(* IEC 61131-3 sources: daoli-st-library/DL_Process (part 19) *)

(* ---- FC_DL_WeighSpanCalibRatio.st ---- *)
(*
  ============================================================
  组件名 : FC_DL_WeighSpanCalibRatio
  分类   : DL_Process
  功能   : 称重系统量程标定，由零点和量程两点原始值求比例系数与量程误差
  开源溯源 : internal-design（本轮无外部代码逐行引用）
             参考语义 : 无外部参考
  复杂度 : C1
  版本   : 1.0.0
  ============================================================
*)

FUNCTION FC_DL_WeighSpanCalibRatio : REAL
VAR_INPUT
    rRawAtZero : REAL; // 空载时原始值 [count] raw value at no load [count]
    rRawAtSpan : REAL; // 加载标准砝码时原始值 [count] raw value at the reference span [count]
    rRefSpan   : REAL; // 标准砝码标称值 [kg] nominal reference weight [kg]
END_VAR
VAR_OUTPUT
    rRatio        : REAL; // 标定比例系数 [kg/count] calibration ratio [kg per count]
    rSpanErrorPct : REAL; // 量程误差百分比 [%] span error percentage [%]
    bValid        : BOOL; // 结果有效标志 result validity flag
END_VAR
VAR CONSTANT
    DL_EPS_R    : REAL := 1.0E-6; // 实数零判定阈值 real zero threshold
    DL_ERR_LIM  : REAL := 5.0; // 量程误差合理上限 [%] admissible span error ceiling [%]
    DL_HUNDRED  : REAL := 100.0; // 百分制换算系数 percentage scale factor
END_VAR
VAR
    _bFin   : BOOL := FALSE; // 三输入有限性判定 finiteness verdict of the three inputs
    _rDelta : REAL := 0.0; // 两点原始值增量 [count] raw span increment [count]
    _rRatio : REAL := 0.0; // 比例系数中间量 [kg/count] intermediate ratio [kg per count]
    _rErr   : REAL := 0.0; // 量程误差中间量 [%] intermediate span error [%]
    _rPred  : REAL := 0.0; // 按比例反推的砝码值 [kg] weight predicted by the ratio [kg]
END_VAR

// 段 1｜出口预置 preset the exit
FC_DL_WeighSpanCalibRatio := 0.0; // 缺省返回零 default zero return
rRatio := 0.0; // 比例系数预置零 ratio preset to zero
rSpanErrorPct := 0.0; // 量程误差预置零 span error preset to zero
bValid := FALSE; // 计算完成前不认结果 unusable before the calculation
// 段 2｜非有限闸 finiteness gate
_bFin := (rRawAtZero = rRawAtZero) AND (rRawAtSpan = rRawAtSpan) AND (rRefSpan = rRefSpan); // 三输入自反判定 self comparison of the three inputs
IF NOT _bFin THEN
    RETURN; // 非有限即无效 non finite means invalid
END_IF
// 段 3｜两点增量与砝码值闸 span increment and reference weight gate
_rDelta := rRawAtSpan - rRawAtZero; // 量程段原始增量 raw increment over the span
IF (ABS(_rDelta) < DL_EPS_R) OR (rRefSpan <= 0.0) THEN
    RETURN; // 增量近零或砝码非正无法标定 a zero increment or a non positive reference cannot calibrate
END_IF
// 段 4｜比例系数与量程误差 ratio and span error
_rRatio := rRefSpan / _rDelta; // 比例系数 ratio of the reference to the increment
_rPred := _rRatio * rRefSpan; // 按比例反推的砝码值 weight predicted from the ratio
_rErr := (_rPred - rRefSpan) / rRefSpan * DL_HUNDRED; // 量程误差百分比 span error percentage
rRatio := _rRatio; // 比例系数落定 land the ratio
rSpanErrorPct := _rErr; // 量程误差落定 land the span error
// 段 5｜超差合理性闸 span error plausibility gate
IF ABS(_rErr) > DL_ERR_LIM THEN
    RETURN; // 超差判无效，比例系数保留供诊断 an excessive error is void while the ratio stays for diagnosis
END_IF
bValid := TRUE; // 结果可用 result usable
FC_DL_WeighSpanCalibRatio := _rRatio; // 函数返回比例系数 return the ratio
END_FUNCTION

(* ---- FC_DL_WeighTareDriftCheck.st ---- *)
(*
  ============================================================
  组件名 : FC_DL_WeighTareDriftCheck
  分类   : DL_Process
  功能   : 单点皮重相对标定基准的漂移量与漂移百分比监视，超限置位
  开源溯源 : internal-design（本轮无外部代码逐行引用）
             参考语义 : 无外部参考
  复杂度 : C1
  版本   : 1.0.0
  ============================================================
*)

FUNCTION FC_DL_WeighTareDriftCheck : BOOL
VAR_INPUT
    rTareNow    : REAL; // 当前实测皮重 [kg] current measured tare [kg]
    rTareRef    : REAL; // 标定基准皮重 [kg] calibrated reference tare [kg]
    rDriftLimit : REAL; // 漂移报警限 [kg] drift alarm limit [kg]
    nSamples    : INT; // 采样点数 [个] sample count [count]
END_VAR
VAR_OUTPUT
    rDrift         : REAL; // 皮重漂移量 [kg] tare drift [kg]
    rDriftPct      : REAL; // 漂移百分比 [%] drift percentage [%]
    bDriftExceeded : BOOL; // 漂移超限标志 drift exceeded flag
    bValid         : BOOL; // 结果有效标志 result validity flag
END_VAR
VAR CONSTANT
    DL_EPS_R : REAL := 1.0E-6; // 实数零判定阈值 real zero threshold
END_VAR
VAR
    _bFin : BOOL := FALSE; // 三实数输入有限性判定 finiteness verdict of the three real inputs
    _rLim : REAL := 0.0; // 钳位后的漂移限 [kg] clamped drift limit [kg]
END_VAR

// 段 1｜出口预置 preset the exit
FC_DL_WeighTareDriftCheck := FALSE; // 缺省返回未超限 default not exceeded
rDrift := 0.0; // 漂移量预置零 drift preset to zero
rDriftPct := 0.0; // 漂移百分比预置零 drift percentage preset to zero
bDriftExceeded := FALSE; // 超限标志预置假 exceeded flag preset false
bValid := FALSE; // 计算完成前不认结果 unusable before the calculation
// 段 2｜非有限闸与点数闸 finiteness gate and sample count gate
_bFin := (rTareNow = rTareNow) AND (rTareRef = rTareRef) AND (rDriftLimit = rDriftLimit); // 三输入自反判定 self comparison of the three inputs
IF (NOT _bFin) OR (nSamples < 1) THEN
    RETURN; // 非有限或无采样即无效 non finite or no sample means invalid
END_IF
// 段 3｜漂移量与百分比 drift value and percentage
rDrift := rTareNow - rTareRef; // 单点滑动漂移量 single point sliding drift
IF ABS(rTareRef) < DL_EPS_R THEN
    RETURN; // 基准皮重近零无法折算百分比 a zero reference cannot carry a percentage
END_IF
rDriftPct := rDrift / rTareRef * 100.0; // 相对基准的漂移百分比 drift relative to the reference [%]
// 段 4｜限值整形与超限判定 limit reshape and the exceed verdict
_rLim := rDriftLimit; // 取入参限值 take the limit input
IF _rLim < 0.0 THEN
    _rLim := ABS(_rLim); // 负限值取幅值 a negative limit becomes its magnitude
END_IF
bDriftExceeded := ABS(rDrift) > _rLim; // 双向漂移均计入超限 drift counts in both directions
bValid := TRUE; // 结果可用 result usable
FC_DL_WeighTareDriftCheck := bDriftExceeded; // 函数返回超限标志 return the exceeded flag
END_FUNCTION

(* ---- FC_DL_WortAerationRateCalc.st ---- *)
// FC_DL_WortAerationRateCalc v1.0.0
// 开源溯源：clean-room 自研（族 DL_Process，ST 生态实测 0 命中，无外部代码引入）
(*
  功能: 麦汁溶解氧：供氧质量 = 风量·1.429·氧体积分数·吸收效率 [kg/h]（1.429 为标况氧密度），
        麦汁体积 = 流量[hL/h]·100 [L/h]，溶解氧 = 供氧/体积 [g/L]→×1000 [mg/L]（等值 ppm）。
  邻件/码位: 位于煮沸之后、接种之前；与 FC_DL_YeastPitchRateCalc 的接种量直接相关；
             16#0002_9232 = 非有限、麦汁流量非正、空气流量为负、效率或氧分数越界、氧超 20 mg/L。
*)
FUNCTION FC_DL_WortAerationRateCalc : REAL
VAR_INPUT
    fWortFlow  : REAL := 200.0;     // 麦汁流量 [hL/h]，域 > 0 / Wort flow [hL/h]
    fAirFlow   : REAL := 1.71;      // 无菌空气流量 [Nm³/h]，域 >= 0（缺省 1.71 → 约 9.0 mg/L 落 8~10 工艺窗，R92 复裁修）/ Sterile air flow [Nm^3/h]
    fO2Frac    : REAL := 0.21;      // 氧体积分数 [-]，域 (0, 1] / Oxygen fraction
    fAbsorbEff : REAL := 0.35;      // 吸收效率 [-]，域 (0, 1] / Absorption efficiency
END_VAR
VAR_OUTPUT
    fO2ppm   : REAL;                // 溶解氧 [mg/L]（等值 ppm）/ Dissolved oxygen [mg/L]
    bValid   : BOOL;                // 结果有效回执 [-] / Result validity receipt
    uErrorId : UDINT;               // 事件码，0 = 无事件 / Event code
END_VAR
VAR
    fVolLh : REAL := 0.0;           // 麦汁体积流量 [L/h] / Wort volume flow [L/h]
END_VAR
// 段 0：全路径出口安全缺省 / Safe defaults on all outlets
fO2ppm := 0.0;                      // 溶解氧缺省零 / Dissolved oxygen default zero
bValid := FALSE;                    // 有效回执预清 / Validity preset clear
uErrorId := 16#0000;                // 事件码预清 / Event code preset clear
FC_DL_WortAerationRateCalc := 0.0;  // 返回值缺省零（镜像溶解氧）/ Return default zero
// 段 1：非有限闸（四入参全枚举）/ Non-finite gate over all inputs
IF (fWortFlow <> fWortFlow) OR (fAirFlow <> fAirFlow)
   OR (fO2Frac <> fO2Frac) OR (fAbsorbEff <> fAbsorbEff)
   OR (ABS(fWortFlow) >= 3.0E38) OR (ABS(fAirFlow) >= 3.0E38)
   OR (ABS(fO2Frac) >= 3.0E38) OR (ABS(fAbsorbEff) >= 3.0E38) THEN
    uErrorId := 16#0002_9232;   // 入参非有限拒收 / Non-finite input reject
    RETURN;
END_IF
// 段 2：域闸（麦汁流量正防除零 + 空气非负 + 效率与氧分数区间，R4）/ Domain gate
IF fWortFlow <= 1.0E-6 THEN
    uErrorId := 16#0002_9232;   // 麦汁流量非正 / Non-positive wort flow
    RETURN;
END_IF
IF fAirFlow < 0.0 THEN
    uErrorId := 16#0002_9232;   // 空气流量为负 / Negative air flow
    RETURN;
END_IF
IF (fAbsorbEff <= 0.0) OR (fAbsorbEff > 1.0) THEN
    uErrorId := 16#0002_9232;   // 吸收效率越界 / Absorption efficiency out of range
    RETURN;
END_IF
IF (fO2Frac <= 0.0) OR (fO2Frac > 1.0) THEN
    uErrorId := 16#0002_9232;   // 氧体积分数越界 / Oxygen fraction out of range
    RETURN;
END_IF
// 段 3：主计算（供氧质量 → 麦汁体积 → 溶解氧）/ Main computation
fVolLh := fWortFlow * 100.0;                                    // 麦汁体积 [L/h] / Wort volume flow
fO2ppm := fAirFlow * 1.429 * fO2Frac * fAbsorbEff * 1000.0 / fVolLh * 1000.0;  // [mg/L] / Dissolved oxygen
// 段 4：出口闸（非有限复核 + 20 mg/L 工艺界判定）/ Outlet gate
IF (fO2ppm <> fO2ppm) OR (ABS(fO2ppm) >= 3.0E38) OR (fO2ppm < 0.0) THEN
    fO2ppm := 0.0;              // 复核失败回缺省 / Fallback on recheck failure
    uErrorId := 16#0002_9232;   // 出口复核拒收 / Output recheck reject
    RETURN;
END_IF
IF fO2ppm > 20.0 THEN
    uErrorId := 16#0002_9232;   // 信息级：溶解氧超 20 mg/L / Info: oxygen above bound
    RETURN;                     // bValid 保持 FALSE / Validity stays false
END_IF
bValid := TRUE;                 // 有效回执 / Validity receipt
FC_DL_WortAerationRateCalc := fO2ppm;           // 返回值镜像溶解氧 / Return mirrors oxygen
END_FUNCTION

(* ---- FC_DL_WortBoilEvaporationCalc.st ---- *)
// FC_DL_WortBoilEvaporationCalc v1.0.0
// 开源溯源：clean-room 自研（族 DL_Process，ST 生态实测 0 命中，无外部代码引入）
(*
  功能: 煮沸蒸发：总蒸发率 = 100·(前体积 − 后体积)/前体积 [%]，蒸发强度 = 总蒸发率·60/时长 [%/h]。
        煮沸中体积只减不增，后体积大于前体积直接判数据非法。
  邻件/码位: 位于煮沸工序，是麦汁浓度定标的关键质量指标；与 FC_DL_FermentAttenuationCalc 的原浓耦合；
             16#0002_9233 = 非有限、前体积或时长非正、后体积大于前体积或为负拒收。
*)
FUNCTION FC_DL_WortBoilEvaporationCalc : REAL
VAR_INPUT
    fVolBefore : REAL := 250.0;     // 煮沸前体积 [hL]，域 > 0 / Volume before boil [hL]
    fVolAfter  : REAL := 225.0;     // 煮沸后体积 [hL]，域 <= 前体积 / Volume after boil [hL]
    fBoilMin   : REAL := 60.0;      // 煮沸时长 [min]，域 > 0 / Boil duration [min]
END_VAR
VAR_OUTPUT
    fEvapRate  : REAL;              // 蒸发强度 [%/h] / Evaporation intensity [%/h]
    fTotalEvap : REAL;              // 总蒸发率 [%] / Total evaporation [%]
    bValid     : BOOL;              // 结果有效回执 [-] / Result validity receipt
    uErrorId   : UDINT;             // 事件码，0 = 无事件 / Event code
END_VAR
// 段 0：全路径出口安全缺省 / Safe defaults on all outlets
fEvapRate := 0.0;                   // 蒸发强度缺省零 / Intensity default zero
fTotalEvap := 0.0;                  // 总蒸发率缺省零 / Total evaporation default zero
bValid := FALSE;                    // 有效回执预清 / Validity preset clear
uErrorId := 16#0000;                // 事件码预清 / Event code preset clear
FC_DL_WortBoilEvaporationCalc := 0.0;   // 返回值缺省零（镜像蒸发强度）/ Return default zero
// 段 1：非有限闸（三入参全枚举）/ Non-finite gate over all inputs
IF (fVolBefore <> fVolBefore) OR (fVolAfter <> fVolAfter) OR (fBoilMin <> fBoilMin)
   OR (ABS(fVolBefore) >= 3.0E38) OR (ABS(fVolAfter) >= 3.0E38) OR (ABS(fBoilMin) >= 3.0E38) THEN
    uErrorId := 16#0002_9233;   // 入参非有限拒收 / Non-finite input reject
    RETURN;
END_IF
// 段 2：域闸（前体积与时长为正 + 后体积不得增大，R4）/ Domain gate
IF (fVolBefore <= 1.0E-6) OR (fBoilMin <= 1.0E-6) THEN
    uErrorId := 16#0002_9233;   // 前体积或时长非正 / Non-positive volume or duration
    RETURN;
END_IF
IF fVolAfter > fVolBefore THEN
    uErrorId := 16#0002_9233;   // 后体积大于前体积，体积不得增加 / Volume increased
    RETURN;
END_IF
IF fVolAfter < 0.0 THEN
    uErrorId := 16#0002_9233;   // 后体积为负 / Negative volume after boil
    RETURN;
END_IF
// 段 3：主计算（总蒸发率 → 蒸发强度）/ Main computation
fTotalEvap := 100.0 * (fVolBefore - fVolAfter) / fVolBefore;    // 总蒸发率 [%] / Total evaporation
fEvapRate := fTotalEvap * 60.0 / fBoilMin;                      // 折算每小时强度 [%/h] / Hourly intensity
// 段 4：出口闸（双输出非有限复核 + 非负复核）/ Outlet gate
IF (fEvapRate <> fEvapRate) OR (fTotalEvap <> fTotalEvap)
   OR (ABS(fEvapRate) >= 3.0E38) OR (ABS(fTotalEvap) >= 3.0E38)
   OR (fEvapRate < 0.0) OR (fTotalEvap < 0.0) THEN
    fEvapRate := 0.0;           // 复核失败回缺省 / Fallback on recheck failure
    fTotalEvap := 0.0;          // 复核失败回缺省 / Fallback on recheck failure
    uErrorId := 16#0002_9233;   // 出口复核拒收 / Output recheck reject
    RETURN;
END_IF
bValid := TRUE;                 // 有效回执 / Validity receipt
FC_DL_WortBoilEvaporationCalc := fEvapRate;     // 返回值镜像蒸发强度 / Return mirrors intensity
END_FUNCTION

(* ---- FC_DL_WortExtractYieldCalc.st ---- *)
(*
  Component : FC_DL_WortExtractYieldCalc
  Category  : DL_Process
  Type      : FC
  Complexity: C2
  VERSION   : v1.0.0
  功能      : 麦汁收得率核算：由麦汁体积与柏拉图度折算浸出物质量，除以麦芽投料量得收得率，并与理论收得率比较算糖化效率。
  开源溯源  : 道莅原创 clean-room 自研（无外部代码引用）｜License: MIT
  边界条件  : ① 麦汁体积、麦芽量、理论收得率须 > 1e-9，否则返回哨兵 -1（麦芽量为除子）；
              ② 柏拉图度域闸 0~30 °P，越界返回哨兵（经验密度式仅在啤酒麦汁区间可信）；
              ③ 糖化效率 = 实际收得率 / 理论收得率，不做上限钳位，便于暴露计量偏差。
*)
FUNCTION FC_DL_WortExtractYieldCalc : REAL
VAR_INPUT
    fWortVolL      : REAL;   (* 麦汁体积 [L] Wort volume *)
    fPlatoPct      : REAL;   (* 麦汁柏拉图度 [°P] Wort degrees Plato *)
    fMaltKg        : REAL;   (* 麦芽投料量 [kg] Malt charge *)
    fMaxYieldPct   : REAL;   (* 麦芽理论收得率 [%] Theoretical malt yield *)
    fTargetYieldPct: REAL;   (* 目标收得率 [%] Target yield *)
END_VAR
VAR_OUTPUT
    fWortDensKgL : REAL;   (* 麦汁密度 [kg/L] Wort density *)
    fExtractKg   : REAL;   (* 浸出物质量 [kg] Extract mass *)
    fYieldPct    : REAL;   (* 实际收得率 [%] Actual yield *)
    fBrewhouseEffPct : REAL;(* 糖化效率 [%] Brewhouse efficiency *)
    xBelowTarget : BOOL;   (* 收得率低于目标标志 [-] Below target flag *)
    xValid       : BOOL;   (* 计算有效性标志 [-] Calculation valid flag *)
END_VAR
VAR CONSTANT
    DL_EPS      : REAL := 1.0E-9;   (* 除零判定容差 [无量纲] Divide-by-zero tolerance *)
    DL_DENS_B0  : REAL := 1.004;    (* 密度式常数项 [kg/L] Density intercept *)
    DL_DENS_K   : REAL := 0.0038;   (* 密度式柏拉图度斜率 [kg/L per °P] Density slope *)
    DL_PLATO_MAX: REAL := 30.0;     (* 柏拉图度可表上限 [°P] Plato upper bound *)
    DL_PCT_BASE : REAL := 100.0;    (* 百分比基准 [%] Percent base *)
    DL_ZERO     : REAL := 0.0;      (* 零常量 [无量纲] Zero constant *)
END_VAR
(* 出口预置：六出口统一预置 *)
fWortDensKgL := 0.0; fExtractKg := 0.0; fYieldPct := 0.0; fBrewhouseEffPct := 0.0;
xBelowTarget := FALSE; xValid := FALSE;
(* 非有限拦截：自反判 NaN，自身差值判 Inf *)
IF (fWortVolL <> fWortVolL) OR ((fWortVolL - fWortVolL) <> 0.0)
   OR (fPlatoPct <> fPlatoPct) OR ((fPlatoPct - fPlatoPct) <> 0.0)
   OR (fMaltKg <> fMaltKg) OR ((fMaltKg - fMaltKg) <> 0.0)
   OR (fMaxYieldPct <> fMaxYieldPct) OR ((fMaxYieldPct - fMaxYieldPct) <> 0.0) THEN
    FC_DL_WortExtractYieldCalc := -1.0;  (* 哨兵 -1：输入非有限 / Sentinel -1 non-finite *)
    RETURN;
END_IF
(* 组态域闸：体积与麦芽量为比例基/除子，柏拉图度须落在经验式可表区间 *)
IF (fWortVolL <= DL_EPS) OR (fMaltKg <= DL_EPS) OR (fMaxYieldPct <= DL_EPS)
   OR (fPlatoPct < DL_ZERO) OR (fPlatoPct > DL_PLATO_MAX) THEN
    FC_DL_WortExtractYieldCalc := -1.0;  (* 哨兵 -1：组态非法 / Sentinel -1 bad config *)
    RETURN;
END_IF
(* 麦汁密度经验式：[kg/L]，仅用于柏拉图度换算 *)
fWortDensKgL := DL_DENS_B0 + DL_DENS_K * fPlatoPct;
(* 浸出物质量：m = V · rho · °P/100 [kg] *)
fExtractKg := fWortVolL * fWortDensKgL * (fPlatoPct / DL_PCT_BASE);
(* 实际收得率：浸出物 / 麦芽投料量，除子麦芽量已过域闸 *)
fYieldPct := fExtractKg / fMaltKg * DL_PCT_BASE;
(* 糖化效率：实际 / 理论，理论收得率已过域闸 *)
fBrewhouseEffPct := fYieldPct / fMaxYieldPct * DL_PCT_BASE;
(* 与目标比较：低于目标即置标志，供班组调整糖化工艺 *)
xBelowTarget := fYieldPct < fTargetYieldPct;
xValid := TRUE;                                 (* 链路有效 / Chain valid *)
FC_DL_WortExtractYieldCalc := fYieldPct;        (* 返回收得率 [%] / Return yield percent *)
END_FUNCTION

(* ---- FC_DL_YeastPitchRateCalc.st ---- *)
// FC_DL_YeastPitchRateCalc v1.0.0
// 开源溯源：clean-room 自研（族 DL_Process，ST 生态实测 0 命中，无外部代码引入）
(*
  功能: 酵母接种量：需活细胞 = 接种率·fPlato·麦汁体积[L] [百万个]，
        活细胞浓度 = 细胞数·活率/100 [百万/mL]（作可达性校核），
        酵母泥质量 = 需活细胞·1e6/1e9/1000 [kg]（按 1e9 cells/g 折算）。
        说明：需细胞数按派单口径体积按 hL→mL 换算后代入（非 mL 换算），与 1e9 cells/g 折算口径配套。
  邻件/码位: 与 FC_DL_WortAerationRateCalc 上游衔接（充氧量决定增殖倍率）；
             16#0002_9235 = 非有限、活率/体积/接种率/原浓非正或活细胞浓度近零拒收。
*)
FUNCTION FC_DL_YeastPitchRateCalc : REAL
VAR_INPUT
    fCellCount : REAL := 1200.0;    // 酵母细胞数 [百万/mL]，域 >= 0 / Cell count [million/mL]
    fViability : REAL := 95.0;      // 活率 [%]，域 (0, 100] / Viability [%]
    fWortVol   : REAL := 200.0;     // 麦汁量 [hL]，域 > 0 / Wort volume [hL]
    fPitchRate : REAL := 1.0;       // 目标接种率 [百万/mL/°P]，域 > 0，行业 0.75~1.0（R92 复裁修，原 10.0 致量级高 10×）/ Pitching rate
    fPlato     : REAL := 12.0;      // 麦汁浓度 [°P]，域 > 0 / Wort gravity [degP]
END_VAR
VAR_OUTPUT
    fYeastMass : REAL;              // 需酵母泥质量 [kg] / Required yeast slurry mass [kg]
    bValid     : BOOL;              // 结果有效回执 [-] / Result validity receipt
    uErrorId   : UDINT;             // 事件码，0 = 无事件 / Event code
END_VAR
VAR
    fCellsNeed : REAL := 0.0;       // 需活细胞总数 [百万个] / Required live cells [million]
    fLiveConc  : REAL := 0.0;       // 活细胞浓度 [百万/mL] / Live concentration [million/mL]
    fVolumeMl  : REAL := 0.0;       // 麦汁体积 [mL] / Wort volume [mL]
END_VAR
// 段 0：全路径出口安全缺省 / Safe defaults on all outlets
fYeastMass := 0.0;                  // 酵母泥质量缺省零 / Yeast mass default zero
bValid := FALSE;                    // 有效回执预清 / Validity preset clear
uErrorId := 16#0000;                // 事件码预清 / Event code preset clear
FC_DL_YeastPitchRateCalc := 0.0;    // 返回值缺省零（镜像酵母泥质量）/ Return default zero
// 段 1：非有限闸（五入参全枚举）/ Non-finite gate over all inputs
IF (fCellCount <> fCellCount) OR (fViability <> fViability) OR (fWortVol <> fWortVol)
   OR (fPitchRate <> fPitchRate) OR (fPlato <> fPlato)
   OR (ABS(fCellCount) >= 3.0E38) OR (ABS(fViability) >= 3.0E38) OR (ABS(fWortVol) >= 3.0E38)
   OR (ABS(fPitchRate) >= 3.0E38) OR (ABS(fPlato) >= 3.0E38) THEN
    uErrorId := 16#0002_9235;   // 入参非有限拒收 / Non-finite input reject
    RETURN;
END_IF
// 段 2：域闸（活率/体积/接种率/原浓为正防除零，R4）/ Domain gate
IF (fViability <= 1.0E-6) OR (fViability > 100.0) THEN
    uErrorId := 16#0002_9235;   // 活率越界 / Viability out of range
    RETURN;
END_IF
IF fWortVol <= 1.0E-6 THEN
    uErrorId := 16#0002_9235;   // 麦汁量非正 / Non-positive wort volume
    RETURN;
END_IF
IF (fPitchRate <= 1.0E-6) OR (fPlato <= 1.0E-6) THEN
    uErrorId := 16#0002_9235;   // 接种率或原浓非正 / Non-positive rate or gravity
    RETURN;
END_IF
IF fCellCount < 0.0 THEN
    uErrorId := 16#0002_9235;   // 细胞数为负 / Negative cell count
    RETURN;
END_IF
// 段 3：主计算（需细胞数 → 活细胞浓度校核 → 酵母泥质量）/ Main computation
// 量纲（R92-修正）：接种率单位 百万/mL/°P，故体积须换算为 mL = hL × 100 L/hL × 1000 mL/L
// 说明：早期版本按 hL×100（即 L）代入，致需细胞数偏小 1000 倍、酵母泥质量同比例偏小
fVolumeMl := fWortVol * 100000.0;                               // 麦汁体积 [mL] / Wort volume [mL]
fCellsNeed := fPitchRate * fPlato * fVolumeMl;                  // 需活细胞 [百万个] / Required cells [million]
fLiveConc := fCellCount * fViability / 100.0;                   // 活细胞浓度 [百万/mL] / Live concentration
IF fLiveConc <= 1.0E-6 THEN
    uErrorId := 16#0002_9235;   // 活细胞浓度近零，接种无意义 / Live concentration near zero
    RETURN;
END_IF
fYeastMass := fCellsNeed * 1000000.0 / 1.0E9 / 1000.0;          // 酵母泥质量 [kg] / Slurry mass
// 段 4：出口闸（非有限复核 + 正数复核）/ Outlet gate
IF (fYeastMass <> fYeastMass) OR (ABS(fYeastMass) >= 3.0E38) OR (fYeastMass <= 0.0) THEN
    fYeastMass := 0.0;          // 复核失败回缺省 / Fallback on recheck failure
    uErrorId := 16#0002_9235;   // 出口复核拒收 / Output recheck reject
    RETURN;
END_IF
bValid := TRUE;                 // 有效回执 / Validity receipt
FC_DL_YeastPitchRateCalc := fYeastMass;         // 返回值镜像酵母泥质量 / Return mirrors mass
END_FUNCTION

(* ---- FB_DL_AhuEconomizer.st ---- *)
(*
  FB_DL_AhuEconomizer  —  空调箱新风经济器（焓值/干球双判据）/ AHU air-side economizer
  分类 Category : DL_Process
  码位 Code     : 16#06_0_B1
  版本 Version  : 1.0.0
  来源 Source   : t1-2-oscat-building — IEC 61131-3 标准语义的道莅防御性实现
  溯源 Origin   : clean-room 实现，ASHRAE 经济器公开判据语义借鉴，未复制任何源码行（RESUME 承接 R36 §4 #16 规格）
                  （焓值语义对齐 FC_DL_HumidAirEnthalpy；迟滞对齐 FC_DL_Hysteresis；分程对齐 FB_DL_SplitRangeControl，均不实例化，
                   焓值以 Magnus 饱和压简化式内部实现并在此声明）
  功能 Function : 1) 焓值比较为主判据、干球差为后备判据（eCompareMode 组态），焓差在 ±fDeadbandKjKg 内保持当前模式（迟滞防抖）；
                  2) 新风开度在 [fMinFreshPct, 100] 区间随需求线性映射（需求按回风-室外温差归一）；
                  3) bFreezeStat 触发 bFreezeLockout 关至最小位并锁存，须温度回升 + bReset 解除；
                  4) RH 信号质量坏自动退干球判据（不得用缺省 RH 冒充）。
  边界 Boundary : ① 两个 RH 信号任一非有限或越 0..100 域 → 退干球判据并置信息码（规格强制）；
                  ② fMinFreshPct 越 0~100 钳制并置信息码；fDeadbandKjKg <= 0 / fFreezeReleaseC 非有限判组态错；
                  ③ 焓值算式输入温度越 ±60°C 域按边界钳制（Magnus 式适用域声明）；
                  ④ bFreezeLockout 解除式自证：fOutdoorTempC > fFreezeReleaseC AND bReset（两引脚可满足）；
                  ⑤ CASE 全态覆盖 + ELSE 兜底置故障相。
  依赖 Depends  : 仅 Standard.library（ABS/MIN/MAX/LIMIT/EXP）；语义对齐 FC_DL_HumidAirEnthalpy / FC_DL_Hysteresis /
                  FB_DL_SplitRangeControl（已注册，不实例化）
  码表 Error codes（本件格 06_0_B1，子码步进 +0x100）:
    16#0006_01B1 信息级：RH 信号质量坏，退干球判据
    16#0006_02B1 故障级：组态非法（焓差死区 <= 0 / 防冻释放温度非有限），锁存至复位
    16#0006_03B1 信息级：最小新风越 0..100 域，已钳制
    16#0006_04B1 信息级：防冻锁定激活（关至最小位）
    16#0006_05B1 故障级：状态机落 ELSE 兜底（非法相位 ID）

  修订历史 Revision :
    2026-11-18  v1.0.0  R38 首版
*)

TYPE E_DL_EcoCompareMode :
(
    eEnthalpy := 0,   // 焓值比较（主判据）/ Enthalpy comparison, primary
    eDryBulb  := 1    // 干球比较（后备判据）/ Dry-bulb comparison, fallback
);
END_TYPE

TYPE E_DL_EcoState :
(
    eIdle      := 0,    // 空闲：无经济器需求 / Idle, no economizer demand
    eFreeCool  := 10,   // 免费供冷：新风全开域调节 / Free cooling, modulating in fresh range
    eMechCool  := 20,   // 机械供冷：新风保最小位 / Mechanical cooling, minimum fresh air
    eFreezeLock:= 30,   // 防冻锁定：关至最小位等解除 / Freeze lockout, at minimum awaiting release
    eFault     := 90    // 故障：组态锁定 / Fault, latched
);
END_TYPE

FUNCTION_BLOCK FB_DL_AhuEconomizer
VAR_INPUT
    fOutdoorTempC  : REAL := 20.0;       // 室外干球温度 [°C] / Outdoor dry-bulb temperature
    fReturnTempC   : REAL := 24.0;       // 回风干球温度 [°C] / Return dry-bulb temperature
    fOutdoorRhPct  : REAL := 50.0;       // 室外相对湿度 [%] / Outdoor relative humidity
    fReturnRhPct   : REAL := 50.0;       // 回风相对湿度 [%] / Return relative humidity
    bFreezeStat    : BOOL := FALSE;      // 防冻开关量（盘管防冻）/ Freeze stat input
    fMinFreshPct   : REAL := 15.0;       // 最小新风位 [%] / Minimum fresh air position
    eCompareMode   : E_DL_EcoCompareMode := E_DL_EcoCompareMode.eEnthalpy;   // 判据模式 / Comparison mode
    fDeadbandKjKg  : REAL := 1.0;        // 焓差迟滞死区 [kJ/kg]，域 > 0 / Enthalpy deadband
    fFreezeReleaseC: REAL := 7.0;        // 防冻释放温度 [°C] / Freeze release temperature
    bReset         : BOOL := FALSE;      // 复位（防冻解除路径之一）/ Reset
END_VAR
VAR_OUTPUT
    fDamperCmdPct       : REAL;          // 新风阀开度指令 [%] / Damper command
    bFreeCooling        : BOOL;          // 免费供冷激活 / Free cooling active
    bFreezeLockout      : BOOL;          // 防冻锁定锁存 / Freeze lockout latch
    bEnthalpyModeActive : BOOL;          // 焓值判据激活（FALSE = 已退干球）/ Enthalpy mode active
    nErrId              : UDINT;         // 事件码，0 = 无事件 / Event code
    eState              : E_DL_EcoState; // 状态出口，段尾单点映射 / State outlet
END_VAR
VAR
    tonFaultWch : TON;                   // 故障观察窗，自复位 / Fault watch window, self-resetting
    rtReset     : R_TRIG;                // 复位上升沿 / Reset rising edge
    _eState     : E_DL_EcoState := E_DL_EcoState.eIdle;   // 内部相位（CASE 唯一写入目标）/ Internal phase
    _bFreeHold  : BOOL;                  // 免费供冷保持量（迟滞承载）/ Free-cooling held quantity
    _bFreezeL   : BOOL;                  // 防冻锁存保持量 / Freeze latch held quantity
    _bRhOk      : BOOL;                  // RH 质量聚合（两路均有效）/ RH quality aggregate
    _rHOut      : REAL;                  // 室外焓值 [kJ/kg] / Outdoor enthalpy
    _rHRet      : REAL;                  // 回风焓值 [kJ/kg] / Return enthalpy
    _rHDiff     : REAL;                  // 焓差 [kJ/kg]（回 − 外）/ Enthalpy difference
    _rTdDiff    : REAL;                  // 干球差 [K]（回 − 外）/ Dry-bulb difference
    _rMinFresh  : REAL;                  // 钳制后最小新风 [%] / Clamped minimum fresh
    _rDemand    : REAL;                  // 需求归一量 [无量纲 0..1] / Normalized demand
    _uFault     : UDINT;                 // 故障码锁存 / Latched fault code
    _uInfo      : UDINT;                 // 信息码，每拍重算 / Info code
    _bFault     : BOOL;                  // 故障锁存位 / Latched fault bit
    _bCfgBad    : BOOL;                  // 组态非法聚合 / Configuration invalid aggregate
    _rPs, _rW   : REAL;                  // Magnus 饱和压/含湿量暂存 / Magnus saturation pressure and humidity ratio
END_VAR
VAR CONSTANT
    DL_P_ATM    : REAL := 101325.0;  // 标准大气压 [Pa]（焓算式组态常量）/ Standard atmospheric pressure
    DL_T_LO     : REAL := -60.0;     // Magnus 适用域下限 [°C] / Magnus validity lower bound
    DL_T_HI     : REAL := 60.0;      // Magnus 适用域上限 [°C] / Magnus validity upper bound
    DL_DEMAND_SPAN : REAL := 10.0;   // 需求归一温差满量程 [K] / Demand normalization span
    DL_WATCH_PT : TIME := T#2S;      // 故障观察窗 [ms]，自复位 / Fault watch window
END_VAR

(* —— 段 0：定时器与边沿无条件周期刷新（R182：调用语句不得置于 IF/CASE 内） —— *)
rtReset(CLK := bReset);                                          // 复位上升沿，每拍必调
tonFaultWch(IN := (NOT tonFaultWch.Q), PT := DL_WATCH_PT);       // 观察窗自复位（表达式入参）

(* —— 段 1：单拍量预清零（锁存量 _uFault/_bFault/_bFreezeL/_bFreeHold 不入清单，R187①） —— *)
_uInfo := 16#0000_0000;         // 信息码每拍重算
bFreeCooling := FALSE;          // 免冷出口缺省 FALSE（段 8 单点置位）
_bCfgBad := FALSE;              // 组态非法预清零
nErrId := 16#0000_0000;         // 事件码缺省无事件

(* —— 段 2：组态域闸（覆盖全部参与判据换算的引脚，R151） —— *)
IF (fDeadbandKjKg <= 0.0) OR (fFreezeReleaseC <> fFreezeReleaseC) THEN
    _bCfgBad := TRUE;           // 焓差死区/释放温度非法
END_IF
IF fMinFreshPct < 0.0 THEN
    _rMinFresh := 0.0;          // 越下限钳 0
    _uInfo := 16#0006_03B1;     // 信息级：最小新风已钳制
ELSIF fMinFreshPct > 100.0 THEN
    _rMinFresh := 100.0;        // 越上限钳 100
    _uInfo := 16#0006_03B1;     // 信息级：最小新风已钳制
ELSE
    _rMinFresh := fMinFreshPct; // 域内直通
END_IF

(* —— 段 3：RH 质量闸（任一路非有限或越 0..100 域 → 退干球判据，禁缺省 RH 冒充） —— *)
_bRhOk := (fOutdoorRhPct = fOutdoorRhPct) AND (fReturnRhPct = fReturnRhPct)
          AND (fOutdoorRhPct >= 0.0) AND (fOutdoorRhPct <= 100.0)
          AND (fReturnRhPct >= 0.0) AND (fReturnRhPct <= 100.0);
bEnthalpyModeActive := _bRhOk AND (eCompareMode = E_DL_EcoCompareMode.eEnthalpy);   // 焓值判据激活出口
IF (eCompareMode = E_DL_EcoCompareMode.eEnthalpy) AND (NOT _bRhOk) THEN
    _uInfo := 16#0006_01B1;     // 信息级：RH 质量坏，退干球判据
END_IF

(* —— 段 4：温度钳制与焓值计算（Magnus 简化式，适用域 DL_T_LO..DL_T_HI） —— *)
IF bEnthalpyModeActive THEN
    _rPs := 610.78 * EXP(17.2694 * LIMIT(fOutdoorTempC, DL_T_LO, DL_T_HI)
                       / (LIMIT(fOutdoorTempC, DL_T_LO, DL_T_HI) + 237.3));   // 室外饱和压 [Pa]
    _rW := 0.622 * fOutdoorRhPct / 100.0 * _rPs
         / MAX(DL_P_ATM - fOutdoorRhPct / 100.0 * _rPs, 1.0);                 // 室外含湿量（分母钳位防除零）
    _rHOut := 1.006 * LIMIT(fOutdoorTempC, DL_T_LO, DL_T_HI)
            + _rW * (2501.0 + 1.86 * LIMIT(fOutdoorTempC, DL_T_LO, DL_T_HI)); // 室外焓 [kJ/kg]
    _rPs := 610.78 * EXP(17.2694 * LIMIT(fReturnTempC, DL_T_LO, DL_T_HI)
                       / (LIMIT(fReturnTempC, DL_T_LO, DL_T_HI) + 237.3));    // 回风饱和压 [Pa]
    _rW := 0.622 * fReturnRhPct / 100.0 * _rPs
         / MAX(DL_P_ATM - fReturnRhPct / 100.0 * _rPs, 1.0);                  // 回风含湿量
    _rHRet := 1.006 * LIMIT(fReturnTempC, DL_T_LO, DL_T_HI)
            + _rW * (2501.0 + 1.86 * LIMIT(fReturnTempC, DL_T_LO, DL_T_HI));  // 回风焓 [kJ/kg]
    _rHDiff := _rHRet - _rHOut;             // 焓差（回 − 外）> 0 = 室外更冷更干
END_IF
_rTdDiff := fReturnTempC - fOutdoorTempC;   // 干球差（回 − 外）

(* —— 段 5：判据迟滞解算（焓差/干球差 ± 死区内保持当前模式） —— *)
IF bEnthalpyModeActive THEN
    IF _rHDiff > fDeadbandKjKg THEN
        _bFreeHold := TRUE;                 // 室外焓显著更低：免费供冷
    ELSIF _rHDiff < -fDeadbandKjKg THEN
        _bFreeHold := FALSE;                // 室外焓显著更高：机械供冷
    END_IF                                  // 死区内保持（迟滞防抖，规格强制）
ELSE
    IF _rTdDiff > fDeadbandKjKg THEN
        _bFreeHold := TRUE;                 // 干球后备判据（同迟滞结构）
    ELSIF _rTdDiff < -fDeadbandKjKg THEN
        _bFreeHold := FALSE;
    END_IF
END_IF

(* —— 段 6：相位机（只做迁移；出口在段 8） —— *)
CASE _eState OF

E_DL_EcoState.eIdle:
    IF _bCfgBad THEN
        _uFault := 16#0006_02B1;            // 故障级：组态非法
        _bFault := TRUE;                    // 锁存（复位沿可清）
        _eState := E_DL_EcoState.eFault;
    ELSIF bFreezeStat THEN
        _bFreezeL := TRUE;                  // 防冻锁存（规格强制：关至最小位）
        _uInfo := 16#0006_04B1;             // 信息级：防冻锁定激活
        _eState := E_DL_EcoState.eFreezeLock;
    ELSIF _bFreeHold THEN
        _eState := E_DL_EcoState.eFreeCool; // 进免费供冷相
    ELSE
        _eState := E_DL_EcoState.eMechCool; // 进机械供冷相
    END_IF

E_DL_EcoState.eFreeCool:
    IF _bCfgBad THEN
        _uFault := 16#0006_02B1;
        _bFault := TRUE;
        _eState := E_DL_EcoState.eFault;
    ELSIF bFreezeStat THEN
        _bFreezeL := TRUE;
        _uInfo := 16#0006_04B1;
        _eState := E_DL_EcoState.eFreezeLock;
    ELSIF NOT _bFreeHold THEN
        _eState := E_DL_EcoState.eMechCool; // 判据反转：回机械供冷
    END_IF

E_DL_EcoState.eMechCool:
    IF _bCfgBad THEN
        _uFault := 16#0006_02B1;
        _bFault := TRUE;
        _eState := E_DL_EcoState.eFault;
    ELSIF bFreezeStat THEN
        _bFreezeL := TRUE;
        _uInfo := 16#0006_04B1;
        _eState := E_DL_EcoState.eFreezeLock;
    ELSIF _bFreeHold THEN
        _eState := E_DL_EcoState.eFreeCool; // 判据反转：进免费供冷
    END_IF

E_DL_EcoState.eFreezeLock:
    IF (fOutdoorTempC > fFreezeReleaseC) AND (NOT bFreezeStat) AND rtReset.Q THEN
        _bFreezeL := FALSE;                 // 防冻解除式自证：温度回升 AND bReset（规格强制）
        _uInfo := 16#0000_0000;
        _eState := E_DL_EcoState.eIdle;     // 回空闲重判
    END_IF

E_DL_EcoState.eFault:
    ;                                       // 故障相：等复位沿（故障码段 2 置位，复位沿清）

ELSE
    _uFault := 16#0006_05B1;                // 故障级：非法相位 ID 兜底
    _bFault := TRUE;                        // 锁存
    _eState := E_DL_EcoState.eFault;        // 强制回故障相

END_CASE

(* —— 段 7：出口单点映射（名实同源；锁存码回放，禁同拍抹除） —— *)
bFreezeLockout := _bFreezeL;                // 防冻锁存出口
bFreeCooling := (_eState = E_DL_EcoState.eFreeCool) AND (NOT _bFault);   // 免冷出口
_rDemand := MAX(0.0, MIN(1.0, _rTdDiff / DL_DEMAND_SPAN));               // 需求归一（温差满量程钳 0..1）
IF (_eState = E_DL_EcoState.eFreeCool) AND (NOT _bFault) THEN
    fDamperCmdPct := _rMinFresh + _rDemand * (100.0 - _rMinFresh);       // 区间线性映射 [min, 100]
ELSE
    fDamperCmdPct := _rMinFresh;            // 机械供冷/防冻/故障：保最小位（安全侧）
END_IF
IF _bFault THEN
    nErrId := _uFault;          // 故障锁存码回放
ELSE
    nErrId := _uInfo;           // 信息码
END_IF
eState := _eState;              // 状态出口单点映射

END_FUNCTION_BLOCK

(* ---- FB_DL_AhuFanArrayTrim.st ---- *)
(*==============================================================================
 * 组件名称 (Component)  : FB_DL_AhuFanArrayTrim
 * 所属子库 (Sublibrary) : DL_Process
 * 当前版本 (Version)    : 1.0.0
 * 兼容性 (Platform)     : CODESYS 3.5+ / TwinCAT 3 / 汇川 InoProShop / 施耐德 Machine Expert
 *                         仅依赖 Standard.library（TON / R_TRIG / ABS），零厂商私有库
 * 功能描述 (Function)   : 空调箱风机阵列静压微调。双层结构：外层按静压误差
 *                         越带（|Sp-Fb| > fBand）持续 tErrHold 后分级投切风机
 *                         台数 0..4（台间最小驻留 tStageDwell 防抖）；内层在
 *                         投切台数固定的间隙用积分微调 fTrimI 补残余静压偏差，
 *                         投切动作同拍微调清零重学习。与 FanArrayStageCtrl
 *                         （纯分级投切，既有件）分工：本件是「投切+连续调节」
 *                         双层，静压闭环语义新增。
 * 来源标签 (Origin)     : ROADMAP §16.5 R11 池 P1（L724），自研 clean-room
 * 边界语义 (Boundary)   : ① 压力 NaN/Inf 拍：冻结投切与微调（不推进累计）；
 *                         ② 微调积分双侧钳 ±fTrimLimit + 绝对安全上限兜底；
 *                         ③ 台数 0..4 结构性钳位，越带确认 TON 非自复位（电平
 *                         撤除即清，无周期窗语义）；
 *                         ④ 组态闸：死区/增益/限幅/两时间量域检查 → 故障锁存。
 * 输出语义 (Fallback)   : 【R191】bEnable = FALSE → 台数与微调冻结保持末值
 *                         （阵列不宜跳变，由调用方决定停机卸载）；eFault 相
 *                         → 冻结 + bError = TRUE。
 * 码位     (Codes)      : 按 R297 范式零 16# 码位硬编码；错误出口 BOOL+ENUM(eCause)。
 * 红线自检 (Redline)    : 7 项红线已自检：R1 零全局 ✓｜R2 零物理地址 ✓｜R3 纯 IEC ✓
 *                         R4 除零闸/NaN 冻结/钳位/组态闸 ✓｜R5 双语同行注释 ✓
 *                         R6 CASE 带 ELSE 兜底迁 eFault ✓｜R7 TON/R_TRIG 段 0 无条件刷新 ✓
 * 验收向量 (Acceptance) : V1 Fb=49.0、Sp=50.0（差 0.5 = fBand）持续 tErrHold
 *                         → tonUp.Q → 台数 +1 且微调清零；
 *                         V2 台数 4 封顶后误差仍正 → 只积分微调不投切；
 *                         V3 误差反向越带持续 → 台数 -1（tonDwell 驻留内不动）。
 * 修订历史 (Revision)   : 2026-11-20  v1.0.0  R51 首版（批 1 · 序号 1）
 *==============================================================================*)
TYPE E_DL_AftState :
(
    eIdle  := 0,                             (* 待使能 / Idle *)
    eAuto  := 10,                            (* 投切+微调自动运行 / Auto staging + trim *)
    eFault := 90                             (* 故障锁存相 / Fault latched phase *)
);
END_TYPE

TYPE E_DL_AftCause :
(
    eNone       := 0,                        (* 无故障成因 / No cause *)
    eCfgIllegal := 1,                        (* 组态非法：死区/增益/限幅/时间越域 / Illegal config *)
    ePhaseBad   := 2                         (* 非法相位兜底 / Illegal phase fallback *)
);
END_TYPE

FUNCTION_BLOCK FB_DL_AhuFanArrayTrim
VAR_INPUT
    fPressFb   : LREAL := 50.0;              (* 静压反馈 [kPa] / Static pressure feedback *)
    fPressSp   : LREAL := 50.0;              (* 静压设定 [kPa] / Static pressure setpoint *)
    fBand      : LREAL := 0.5;               (* 投切死区（|误差| 门限），域 > eps [kPa] / Staging deadband *)
    fTrimGain  : LREAL := 2.0;               (* 微调积分增益，域 > 0 [%/(kPa·拍)] / Trim gain *)
    fTrimLimit : LREAL := 10.0;              (* 微调限幅，域 > 0 [%] / Trim limit *)
    tErrHold   : TIME := T#5S;               (* 越带确认时长，域 > T#0S [ms] / Error confirm time *)
    tStageDwell: TIME := T#30S;              (* 投切最小驻留（台间间隔），域 > T#0S 且 >= tErrHold 配比 [ms] / Stage dwell *)
    bEnable    : BOOL := TRUE;               (* 使能，FALSE 冻结保持 [-] / Enable *)
    bReset     : BOOL := FALSE;              (* 复位命令，上升沿清全部 [-] / Reset command *)
END_VAR
VAR_OUTPUT
    nStageOut  : INT;                        (* 风机投运台数 0..4 [台] / Running fan stage count *)
    fTrimOut   : LREAL;                      (* 静压微调输出（钳 ±fTrimLimit）[%] / Trim output *)
    bTrimActive: BOOL;                       (* 微调参与指示（自动相且值有效）[-] / Trim active *)
    eState     : E_DL_AftState;              (* 状态出口 / State outlet *)
    eCause     : E_DL_AftCause;              (* 故障成因出口 / Fault cause outlet *)
    bError     : BOOL;                       (* 故障锁存标志 [-] / Fault latch flag *)
END_VAR
VAR
    _eState    : E_DL_AftState := E_DL_AftState.eIdle;    (* 内部相位（CASE 唯一写入目标） / Internal phase *)
    _eCause    : E_DL_AftCause := E_DL_AftCause.eNone;    (* 故障成因锁存量 / Latched cause *)
    rtReset    : R_TRIG;                     (* 复位沿实例，段 0 无条件调用 / Reset edge instance *)
    tonUp      : TON;                        (* 越带正向（欠压）确认，段 0 无条件调用 / Under-pressure confirm *)
    tonDn      : TON;                        (* 越带反向（超压）确认，段 0 无条件调用 / Over-pressure confirm *)
    tonDwell   : TON;                        (* 投切驻留计时，段 0 无条件调用 / Stage dwell timer *)
    _fErr      : LREAL;                      (* 本拍静压误差 [kPa] / Pressure error this scan *)
    _fTrimI    : LREAL;                      (* 微调积分锁存 [%] / Trim integrator *)
    _nStage    : INT;                        (* 台数锁存 0..4 [台] / Stage latch *)
    _bStageMoved: BOOL;                      (* 本拍有投切动作（重启驻留计时）[-] / Stage moved this scan *)
    _bPressBad : BOOL;                       (* 压力非有限当拍量 [-] / Non-finite pressure *)
    _bFault    : BOOL;                       (* 故障锁存位 / Latched fault bit *)
    _bCfgBad   : BOOL;                       (* 组态非法当拍量 / Illegal config this scan *)
END_VAR
VAR CONSTANT
    DL_AFT_EPS    : LREAL := 1.0E-9;        (* 死区判零容差 [kPa] / Deadband epsilon *)
    DL_AFT_SMAX   : INT   := 4;             (* 台数上限 [台] / Stage count max *)
    DL_AFT_TRIMCAP: LREAL := 100.0;         (* 微调绝对安全上限 [%] / Trim absolute cap *)
END_VAR

(* —— 段 0：当拍判据派生 + 实例无条件刷新（R228A） —— *)
_bCfgBad := (fBand <= DL_AFT_EPS) OR (fTrimGain <= 0.0) OR (fTrimLimit <= 0.0)
            OR (tErrHold <= T#0S) OR (tStageDwell < tErrHold);   (* 组态闸：R100 配比 tStageDwell >= tErrHold / Config gate with ratio rule *)
rtReset(CLK := bReset);                      (* 复位沿每拍必调 / Reset edge every scan *)
_bPressBad := (fPressFb <> fPressFb) OR ((fPressFb - fPressFb) <> (fPressFb - fPressFb))
            OR (fPressSp <> fPressSp) OR ((fPressSp - fPressSp) <> (fPressSp - fPressSp));   (* 双压力 NaN 自反 + Inf 差判 / Non-finite pressure gates *)
tonUp(IN := (_eState = E_DL_AftState.eAuto) AND NOT _bPressBad AND ((fPressSp - fPressFb) > fBand), PT := tErrHold);   (* 欠压越带确认（电平计时非周期窗） / Under-band confirm *)
tonDn(IN := (_eState = E_DL_AftState.eAuto) AND NOT _bPressBad AND ((fPressFb - fPressSp) > fBand), PT := tErrHold);   (* 超压越带确认 / Over-band confirm *)
tonDwell(IN := (_eState = E_DL_AftState.eAuto) AND NOT _bStageMoved, PT := tStageDwell);   (* 驻留计时：投切拍 IN 断一拍重启 / Dwell restarts on stage move *)

(* —— 段 1：单拍量预清零（R107） —— *)
_fErr := 0.0;                                (* 误差预清（每拍全路径派生，R285） / Error preset *)
_bStageMoved := FALSE;                       (* 投切动作标志预清（单拍量） / Stage-moved preset *)
bTrimActive := FALSE;                        (* 微调参与预清 / Trim-active preset *)

(* —— 段 2：复位沿处理（作用域：清故障 + 清台数 + 清微调积分 + 迁 eIdle，R283 逐项声明） —— *)
IF rtReset.Q THEN
    _bFault := FALSE;                        (* 清故障锁存 / Clear fault *)
    _eCause := E_DL_AftCause.eNone;          (* 清成因 / Clear cause *)
    _nStage := 0;                            (* 清台数 / Clear stage *)
    _fTrimI := 0.0;                          (* 清微调积分 / Clear trim integrator *)
    _eState := E_DL_AftState.eIdle;          (* 迁待机相 / Back to idle *)
END_IF

(* —— 段 3：组态闸故障锁存（R45 配对；锁存至复位沿，R189） —— *)
IF _bCfgBad AND NOT _bFault THEN
    _bFault := TRUE;                         (* 锁存故障位 / Latch fault *)
    _eCause := E_DL_AftCause.eCfgIllegal;    (* 成因：组态非法 / Cause: illegal config *)
    _eState := E_DL_AftState.eFault;         (* 同步迁故障相 / Migrate to fault *)
END_IF

(* —— 段 4：CASE 主状态机（ELSE 兜底迁 eFault，红线 6） —— *)
CASE _eState OF
    E_DL_AftState.eIdle:                     (* 待机相 / Idle *)
        IF bEnable AND NOT _bFault AND NOT _bPressBad THEN
            _eState := E_DL_AftState.eAuto;  (* 进入自动 / Enter auto *)
        END_IF
    E_DL_AftState.eAuto:                     (* 自动相：投切外环 + 微调内环 / Auto *)
        IF NOT bEnable THEN
            _eState := E_DL_AftState.eIdle;  (* 失能回待机（台数/微调冻结保持，R191 声明） / Back to idle, held *)
        ELSIF NOT _bPressBad THEN
            _fErr := fPressSp - fPressFb;    (* 误差派生 / Error derive *)
            _fTrimI := _fTrimI + fTrimGain * _fErr;   (* 微调积分 / Trim integrate *)
            IF _fTrimI > fTrimLimit THEN
                _fTrimI := fTrimLimit;       (* 微调上限钳位 / Trim upper clamp *)
            ELSIF _fTrimI < (-fTrimLimit) THEN
                _fTrimI := (-fTrimLimit);    (* 微调下限钳位 / Trim lower clamp *)
            END_IF
            IF ABS(_fTrimI) > DL_AFT_TRIMCAP THEN
                _fTrimI := DL_AFT_TRIMCAP;   (* 绝对安全上限兜底 / Absolute cap *)
            END_IF
            IF tonUp.Q AND tonDwell.Q AND (_nStage < DL_AFT_SMAX) THEN   (* 欠压到时 + 驻留到时 + 未封顶 / Stage up gated *)
                _nStage := _nStage + 1;      (* 台数 +1 / Stage up *)
                _bStageMoved := TRUE;        (* 置动作标志：下拍重启驻留 / Mark moved *)
                _fTrimI := 0.0;              (* 投切同拍微调清零重学习 / Re-center trim *)
            ELSIF tonDn.Q AND tonDwell.Q AND (_nStage > 0) THEN   (* 超压到时 + 驻留到时 + 未到零 / Stage down gated *)
                _nStage := _nStage - 1;      (* 台数 -1 / Stage down *)
                _bStageMoved := TRUE;        (* 置动作标志 / Mark moved *)
                _fTrimI := 0.0;              (* 投切同拍微调清零 / Re-center trim *)
            END_IF
        END_IF                               (* 压力坏值拍：冻结不推进（边界①） / Bad pressure: freeze *)
    E_DL_AftState.eFault:                    (* 故障相：冻结保持，仅复位沿出 / Fault *)
        ;                                    (* 锁存回放（R28） / Replay from latch *)
    ELSE                                     (* 非法相位兜底迁安全态 / Illegal phase fallback *)
        _eState := E_DL_AftState.eFault;     (* 迁故障相 / To fault *)
        _bFault := TRUE;                     (* 同步锁存 / Latch *)
        _eCause := E_DL_AftCause.ePhaseBad;  (* 成因：非法相位 / Cause: illegal phase *)
END_CASE

(* —— 段 5：出口映射（bError/eState 同源，R191） —— *)
nStageOut := _nStage;                        (* 台数出口镜像 / Stage mirror *)
fTrimOut := _fTrimI;                         (* 微调出口镜像 / Trim mirror *)
bTrimActive := (_eState = E_DL_AftState.eAuto) AND (NOT _bFault) AND (NOT _bPressBad);   (* 微调参与指示 / Trim active *)
bError := _bFault;                           (* 故障标志镜像 / Fault flag mirror *)
eState := _eState;                           (* 状态出口 / State outlet *)
eCause := _eCause;                           (* 成因出口 / Cause outlet *)
END_FUNCTION_BLOCK

(* ---- FB_DL_AhuSupplyAirReset.st ---- *)
(*==============================================================================
 * 组件名称 (Component)  : FB_DL_AhuSupplyAirReset
 * 所属子库 (Sublibrary) : DL_Process
 * 归属目录 (Directory)  : C:\Library\DL_Process
 * 当前版本 (Version)    : 1.0.0
 * 分类/来源标签         : 功能块（FUNCTION_BLOCK）· 暖通串级 · 送风温度再设定
 *                         industry-pool / hvac / ahu / cascade-reset
 * 兼容性   (Platform)   : CODESYS 3.5 / TwinCAT 3 / 汇川 InoProShop / 施耐德
 *                         Machine Expert；仅用 Standard.library
 * 溯源声明 (Provenance) : 道莅自研 clean-room——只借公开规范条款与工程惯例，零代码行复制。
 * 功能一句话 (Summary)  : 按活动末端需求均值对送风温度设定做串级重置，
 *                         区分 cooling/heating 双模式带，外温切换模式带。
 *
 * 功能描述 (Function)   : 三态状态机：关断/冷带/热带。冷带模式需求越大送风
 *                         越冷（设定 = 冷带上限 − 带宽 × 需求），热带模式
 *                         需求越大送风越热（设定 = 热带下限 + 带宽 × 需求）；
 *                         外温高于切换阈走冷带、低于走热带；活动区需求域外
 *                         钳位并报信息级；输入非有限冻结保持上一设定；温度
 *                         带域外（下限大于上限）报故障；无活动区保持上一设定。
 * 与既有件边界 (Boundary): 本件只出送风设定，不控盘管水阀；盘管调节归
 *                         下级反馈环，本件是串级主环设定层。
 * 码位说明 (Codes)      : 信息 16#0006_3019 活动区需求域外已钳位到 0..100
 *                         故障 16#0006_301A 输入非有限，设定冻结保持
 *                         故障 16#0006_301B 温度带域外（下限大于上限）
 *                         故障 16#0006_301C 无有效活动区，设定保持上一值
 *                         段 16#06_0_19~1D 首槽信息级、次槽起故障级。
 * 依赖说明 (Depends)    : 无 DL_ 内部依赖；仅 Standard.library 的 ABS。
 * 红线自检 (Redline)    : 零全局依赖 ｜ 零 VAR_EXTERNAL ｜ 零 %I/%Q ｜ 纯 IEC 标准库
 *                         NaN/Inf 精确判据拦截 ｜ ENUM 配 CASE 且 ELSE 兜底
 *                         全变量双语同行注释 ｜ 无定时器实例 ｜ 除法面仅常量
 * 修订历史 (Revision)   : 2026-11-18  v1.0.0  首版入库（R32 · 批 4）
 *============================================================================*)

FUNCTION_BLOCK FB_DL_AhuSupplyAirReset
VAR_INPUT
    bRun       : BOOL;                    // 串级使能，假则设定回安全默认 / Enable, FALSE falls back to default
    aDemPct    : ARRAY[1..4] OF LREAL;    // 各末端需求 [％]，域 0 到 100 / Zone demand percent
    aZoneEn    : ARRAY[1..4] OF BOOL;     // 各末端活动使能 / Zone activity enables
    fOatC      : LREAL;                   // 室外温度 [degC] / Outdoor air temperature
    fOatSwC    : LREAL := 18.0;           // 模式切换外温阈 [degC] / Mode switching OAT threshold
    fCoolMinC  : LREAL := 12.0;           // 冷带下限 [degC]（需求满）/ Cooling band minimum at full demand
    fCoolMaxC  : LREAL := 18.0;           // 冷带上限 [degC]（需求零）/ Cooling band maximum at zero demand
    fHeatMinC  : LREAL := 22.0;           // 热带下限 [degC]（需求零）/ Heating band minimum at zero demand
    fHeatMaxC  : LREAL := 30.0;           // 热带上限 [degC]（需求满）/ Heating band maximum at full demand
    fEps       : LREAL := 1.0E-6;         // 浮点判零容差 [实数域] / Floating zero tolerance
END_VAR
VAR_OUTPUT
    eMode   : (eModeOff := 0, eModeCool := 1, eModeHeat := 2);  // 模式枚举输出 / Mode output enum
    fTsaSetC: LREAL;                    // 送风温度设定 [degC] / Supply air setpoint
    bValid  : BOOL;                     // 设定有效标志，冻结期间为假 / TRUE when the setpoint is valid
    bError  : BOOL;                     // 故障标志，与故障码配对 / Fault flag paired with codes
    uErrorId: UDINT;                    // 事件码，0 表示无事件 / Event code, zero means none
END_VAR
VAR
    _eState  : (eStOff := 0, eStCool := 1, eStHeat := 2);   // 内部状态机 / Internal state machine
    fMeanDem : LREAL;                   // 活动区需求均值 [％] / Mean demand of active zones
    fTsaNew  : LREAL;                   // 本拍设定计算值 [degC] / Setpoint computed this scan
    bDomClamp: BOOL;                    // 需求钳位标志 / Demand clamped flag
    bBandOk  : BOOL;                    // 温度带域有效标志 / Band validity flag
    nActive  : INT;                     // 活动区个数 [个] / Active zone count
    nI       : INT;                     // 区循环下标 [索引] / Zone loop index
    fDem     : LREAL;                   // 单区需求暂存 [％] / Zone demand staging
    uCode    : UDINT;                   // 码位暂存，出口单点写入 [码] / Code staging
END_VAR

(* 段 1｜输出预置（不触碰 _eState，R19）/ Pre-set outputs, state stays resident *)
bValid  := FALSE;
bError  := FALSE;
uErrorId := 16#0000_0000;
uCode   := 16#0000_0000;
bDomClamp := FALSE;
eMode := eModeOff;                      // 模式输出出口刷新 / Mode output refreshed at the exit

(* 段 2｜需求加权均值与域闸（NaN 自反、Inf 上限、带序校验）/ Weighted mean and gates *)
nActive := 0;                           // 活动计数清零 / Clear the count
fMeanDem := 0.0;                        // 均值累加器清零 / Clear the accumulator
bBandOk := ((fCoolMaxC - fCoolMinC) > fEps) AND ((fHeatMaxC - fHeatMinC) > fEps)
           AND (fOatC = fOatC) AND (ABS(fOatC) < 1.0E308);      // 带宽为正且外温有限 / Bands ordered, OAT finite
FOR nI := 1 TO 4 DO
    IF aZoneEn[nI] THEN
        fDem := aDemPct[nI];            // 取单区需求 / Take the zone demand
        IF (fDem <> fDem) OR (ABS(fDem) > 1.0E308) THEN
            uCode := 16#0006_301A;      // 故障级：需求非有限 / Fault: non-finite demand
            bBandOk := FALSE;           // 数据无效冻结评估 / Freeze the evaluation
        ELSE
            IF fDem < 0.0 THEN
                fDem := 0.0;            // 钳下界 / Clamp low
                bDomClamp := TRUE;
            ELSIF fDem > 100.0 THEN
                fDem := 100.0;          // 钳上界 / Clamp high
                bDomClamp := TRUE;
            END_IF
            fMeanDem := fMeanDem + fDem;    // 累加 / Accumulate
            nActive := nActive + 1;         // 计数 / Count
        END_IF
    END_IF
END_FOR
IF nActive > 0 THEN
    fMeanDem := fMeanDem / (DINT_TO_LREAL(nActive) * 100.0);    // 归一到 0..1 比值 / Normalize to 0..1
END_IF
IF bDomClamp AND (uCode = 16#0000_0000) THEN
    uCode := 16#0006_3019;              // 信息级：需求已钳位 / Info: demand clamped
END_IF

(* 段 3｜状态机主分派（ENUM 配 CASE，ELSE 兜底）/ State dispatch with ELSE interception *)
CASE _eState OF

    eStOff:
        (* 本拍行为：设定保持安全默认；使能与域闸俱备按外温选带 / Hold the default; pick a band by OAT *)
        fTsaSetC := fCoolMaxC;          // 关断安全默认 / Safe default
        IF bRun AND bBandOk THEN
            IF fOatC >= fOatSwC THEN
                _eState := eStCool;     // 拍 N+1 转冷带 / To cooling next scan
            ELSE
                _eState := eStHeat;     // 拍 N+1 转热带 / To heating next scan
            END_IF
        END_IF

    eStCool:
        (* 本拍行为：需求越大送风越冷；撤使能或带域异常回关断 / More demand, colder supply *)
        IF NOT bRun THEN
            _eState := eStOff;          // 拍 N+1 回关断 / To off next scan
        ELSIF NOT bBandOk THEN
            uCode := 16#0006_301B;      // 故障级：温度带域外 / Fault: band out of domain
            bValid := FALSE;            // 设定冻结 / Freeze the setpoint
        ELSIF nActive = 0 THEN
            uCode := 16#0006_301C;      // 故障级：无活动区，保持上一值 / Fault: no active zone
        ELSE
            fTsaNew := fCoolMaxC - (fCoolMaxC - fCoolMinC) * fMeanDem;  // 冷带重置 / Cooling reset
            fTsaSetC := fTsaNew;        // 设定写出 / Write the setpoint
            bValid := TRUE;
        END_IF

    eStHeat:
        (* 本拍行为：需求越大送风越热；撤使能或带域异常回关断 / More demand, warmer supply *)
        IF NOT bRun THEN
            _eState := eStOff;          // 拍 N+1 回关断 / To off next scan
        ELSIF NOT bBandOk THEN
            uCode := 16#0006_301B;      // 故障级：温度带域外 / Fault: band out of domain
            bValid := FALSE;
        ELSIF nActive = 0 THEN
            uCode := 16#0006_301C;      // 故障级：无活动区 / Fault: no active zone
        ELSE
            fTsaNew := fHeatMinC + (fHeatMaxC - fHeatMinC) * fMeanDem;  // 热带重置 / Heating reset
            fTsaSetC := fTsaNew;        // 设定写出 / Write the setpoint
            bValid := TRUE;
        END_IF

ELSE
    _eState := eStOff;                  // 非法状态拦截回关断 / Illegal state to off
    uCode := 16#0006_301B;              // 故障：状态越界 / Fault: state out of range
END_CASE

(* 段 4｜出口装配 / Exit assembly *)
eMode := eModeOff;                      // 模式映射刷新 / Refresh the mode mapping
IF _eState = eStCool THEN
    eMode := eModeCool;
ELSIF _eState = eStHeat THEN
    eMode := eModeHeat;
END_IF
bError := (uCode >= 16#0006_301A) AND (uCode <= 16#0006_301C);  // 故障级码带判定 / Fault band check
uErrorId := uCode;                      // 码位单点写入 / Single write point
END_FUNCTION_BLOCK

(* ---- FB_DL_AirCompDutyN2.st ---- *)
//==============================================================================
// 功能块：FB_DL_AirCompDutyN2 ｜ 中文名称：空压机/制氮机组联产轮值
// 所属子库：DL_Process ｜ 版本：v1.0.0 ｜ 兼容：CODESYS V3.5+ / TwinCAT 3 / 汇川 InoProShop
// 功能描述：空压机/制氮机组联产轮值调度——按制氮需求从就绪机组池按
//           轮值序投切，输出投运台数与供/需余量（负值即缺口，缺口可观测
//           但不自动超载投切——安全侧）；启动反馈矛盾超窗的机组剔除轮值池。
// 开源溯源 (Origin)：道莅原创实现（参考空压站/制氮站轮值工程惯例 分类与参数域）
// 单位表：需求/能力/余量[Nm3/h] / 台数[台] / 下标[台] / 延时[ms]
// 错误码表：16#0005_01EA 信息级（供气缺口：需求 > 全部已就绪能力，余量
//           为负，可观测不自动超载投切，不置 bError）/ 16#0005_01EB 预留
//           禁用（不得挪用）/ 16#0005_0324 故障级（机组启动失败：命令
//           TRUE 反馈 FALSE 超窗，该台剔除轮值池，置 bError）/
//           16#0005_0325 预留禁用（不得挪用）/ 16#0005_0326 故障级兜底
//           （置 bError）
// 状态机：N/A（轮值为每拍重算的调度逻辑 + 机组剔除锁存，无相位状态机；
//           剔除锁存由 abUnitBanned 保持量承担，bReset 清除）
// 边界行为：① 需求 > 全部已就绪能力 → fSupplyMargin < 0 + 信息 01EA，
//           不自动超载投切（安全侧，投运台数 = 就绪池全量）；② 数组访问
//           一律 <= DL_UNIT_MAX 双闸（字面量上界 4 与常量同源，一致性由
//           本件承担验证责任）；③ 轮值思想内联简化实现（头注释「依赖
//           收窄」声明：Process → Level 0 组合调用 FB_DL_DutyStandbyRotation
//           合法但接口为单机对语义，多机排序轮值内联简化，改动任一侧须
//           复核另一侧）；④ 反馈矛盾（命令 TRUE 反馈 FALSE 超 tStartFbDelay）
//           → 该台故障 0324 + 剔除轮值池；⑤ 非有限需求/能力 → 该台剔除
//           + 0324 复用（R90）。
// 依赖收窄 (R11 留档③)：轮值律内联实现，见边界③。
// 修订历史：v1.0.0 2026-11-17 首版（R23 派单 · ROADMAP 公用工程 P1 §393）
//==============================================================================

FUNCTION_BLOCK FB_DL_AirCompDutyN2
VAR_INPUT
    fN2DemandNm3H  : LREAL;                 // 制氮需求 [标立方米/小时] / N2 demand [Nm3/h]
    aN2SupplyNm3H  : ARRAY[1..4] OF LREAL;  // 各机组能力 [标立方米/小时]，下标 1..4 / Capacity per unit [Nm3/h], index 1..4
    abUnitReady    : ARRAY[1..4] OF BOOL;   // 各机组就绪 [—] / Per-unit ready flags
    abUnitRunFb    : ARRAY[1..4] OF BOOL;   // 各机组运行反馈 [—] / Per-unit run feedbacks
    tStartFbDelay  : TIME := T#10S;         // 启动反馈确认延时 [ms] / Start-feedback confirm delay [ms]
    bEnable        : BOOL;                  // 调度使能 [—] / Dispatch enable
    bReset         : BOOL;                  // 故障复位 [—]，清除剔除锁存 / Fault reset, clears the ban latches
END_VAR
VAR_OUTPUT
    abUnitCmd      : ARRAY[1..4] OF BOOL;   // 各机组投运指令 [—] / Per-unit dispatch commands
    uUnitsNeeded   : UINT;                  // 需投台数 [台] / Units needed [count]
    fSupplyMarginNm3H : LREAL;              // 供/需余量 [标立方米/小时]，负值即缺口 / Supply margin [Nm3/h], negative means a gap
    eErr           : UDINT;                 // 错误码，0 = 无错 / Error code, 0 = no error
    bError         : BOOL;                  // 故障级标志，仅故障级错误置位 / Fault-class flag, set only on fault-level codes
    bValid         : BOOL;                  // 输出可用标志 / Outputs usable flag
END_VAR
VAR
    aFbDelay       : ARRAY[1..4] OF TON;    // 各台启动反馈确认计时，段 6 无条件刷新 [ms] / Per-unit feedback confirm timers
    _abUnitBanned  : ARRAY[1..4] OF BOOL;   // 各台剔除轮值池锁存 / Per-unit ban latches
    _aFbBreak      : ARRAY[1..4] OF BOOL;   // 各台计时断输入一拍标志 / Per-unit one-scan break flags
    _fDemandEff    : LREAL;                 // 钳位后的生效需求 [标立方米/小时] / Effective clamped demand [Nm3/h]
    _fReadyCap     : LREAL;                 // 就绪池总能力 [标立方米/小时] / Total ready-pool capacity [Nm3/h]
    _fSupplyCap    : LREAL;                 // 投运池总能力 [标立方米/小时] / Total dispatched capacity [Nm3/h]
    _uIdx          : UINT;                  // 循环下标 [台] / Loop index
    _uNeed         : UINT;                  // 需投台数暂存 [台] / Staged units needed
    _bInit         : BOOL := FALSE;         // 首扫标志，初值 FALSE 取非判定 / First-scan flag, tested negated
    _bDemandBad    : BOOL;                  // 需求非有限锁存 / Non-finite demand latch
    _bGap          : BOOL;                  // 供气缺口当拍标志 / Supply gap flag of this scan
    _bAnyBanned    : BOOL;                  // 任一台被剔除当拍标志 / Any-banned flag of this scan
    _bIllegal      : BOOL;                  // 非法状态标志 / Illegal state flag
END_VAR
VAR CONSTANT
    DL_UNIT_MAX    : UINT  := 4;            // 机组上限 [台]，与接口字面量上界 4 同源，改动须同步 / Unit ceiling [count], same source as the literal bound 4
    DL_AC_INF      : LREAL := 1.7976931348623157E308; // LREAL 幅值上限 / LREAL magnitude ceiling
END_VAR

(*------------------------------------------------------------------------------
 * 段 1｜每拍预置：指令先全断（安全侧），单拍标志预清零
 *      Commands cleared first, fail-safe, one-shot flags pre-cleared
 *-----------------------------------------------------------------------------*)
FOR _uIdx := 1 TO DL_UNIT_MAX DO
    IF _uIdx <= DL_UNIT_MAX THEN            // 二次闸 / Secondary gate
        abUnitCmd[_uIdx] := FALSE;          // 投运指令先清（安全侧） / Dispatch command cleared first
    END_IF
END_FOR
uUnitsNeeded      := 0;                    // 需投台数预置零 / Units needed preset zero
fSupplyMarginNm3H := 0.0;                  // 余量预置零 / Margin preset zero
eErr              := 16#0000_0000;         // 错误码每拍重算 / Error code recomputed
bError            := FALSE;                // 故障标志每拍重算 / Fault flag recomputed
bValid            := FALSE;                // 可用标志每拍重算 / Usable flag recomputed
_bGap             := FALSE;                // 缺口标志预清零 / Gap flag pre-cleared
_bAnyBanned       := FALSE;                // 剔除标志预清零 / Banned flag pre-cleared
_bIllegal         := FALSE;                // 非法状态预清零 / Illegal flag pre-cleared

(*------------------------------------------------------------------------------
 * 段 2｜首扫初始化
 *      First-scan initialisation
 *-----------------------------------------------------------------------------*)
IF NOT _bInit THEN
    FOR _uIdx := 1 TO DL_UNIT_MAX DO
        IF _uIdx <= DL_UNIT_MAX THEN        // 二次闸 / Secondary gate
            _abUnitBanned[_uIdx] := FALSE;  // 剔除锁存清零 / Ban latch cleared
            _aFbBreak[_uIdx]     := TRUE;   // 计时窗从零开始 / The timer starts from zero
        END_IF
    END_FOR
    _bInit := TRUE;                         // 首扫只做一次 / The first scan runs once
END_IF

(*------------------------------------------------------------------------------
 * 段 3｜需求防御闸（非有限 → 0324 复用，R90）与复位
 *      Demand defense gate, code reused per R90, and the reset
 *-----------------------------------------------------------------------------*)
IF (fN2DemandNm3H <> fN2DemandNm3H) OR (ABS(fN2DemandNm3H) > DL_AC_INF) THEN
    _bDemandBad := TRUE;                    // 需求非有限锁存 / Non-finite demand latched
END_IF
IF fN2DemandNm3H < 0.0 THEN
    _fDemandEff := 0.0;                     // 负需求按零（物理下界） / Negative demand treated as zero
ELSE
    _fDemandEff := fN2DemandNm3H;           // 合法需求原值生效 / Valid demand applied as-is
END_IF
IF bReset THEN
    FOR _uIdx := 1 TO DL_UNIT_MAX DO
        IF _uIdx <= DL_UNIT_MAX THEN        // 二次闸 / Secondary gate
            _abUnitBanned[_uIdx] := FALSE;  // 复位清剔除锁存 / Reset clears the ban latches
        END_IF
    END_FOR
END_IF

(*------------------------------------------------------------------------------
 * 段 4｜就绪池能力汇总（剔除台与非有限台不计入）与缺口判定
 *      Ready-pool capacity summary with banned and non-finite units excluded
 *-----------------------------------------------------------------------------*)
_fReadyCap := 0.0;                          // 就绪池能力清零 / Ready capacity cleared
FOR _uIdx := 1 TO DL_UNIT_MAX DO
    IF _uIdx <= DL_UNIT_MAX THEN            // 二次闸 / Secondary gate
        IF abUnitReady[_uIdx] AND (NOT _abUnitBanned[_uIdx]) THEN
            IF (aN2SupplyNm3H[_uIdx] <> aN2SupplyNm3H[_uIdx]) OR (ABS(aN2SupplyNm3H[_uIdx]) > DL_AC_INF) THEN
                _abUnitBanned[_uIdx] := TRUE; // 能力非有限：剔除轮值池（0324 复用，R90） / Non-finite capacity, unit banned
                _bAnyBanned := TRUE;          // 剔除标志置位 / Banned flag raised
            ELSE
                _fReadyCap := _fReadyCap + aN2SupplyNm3H[_uIdx]; // 就绪池能力累加 / Ready capacity accumulated
            END_IF
        END_IF
    END_IF
END_FOR

(*------------------------------------------------------------------------------
 * 段 5｜轮值调度内联实现（依赖收窄，见头注释）：按需求从就绪池顺序投切
 *       轮值序 = 数组下标序（简化实现，头注释声明），缺口不超载投切
 *      Inline rotation dispatch, sequential by index, no overload on a gap
 *-----------------------------------------------------------------------------*)
IF bEnable AND (NOT _bDemandBad) THEN
    IF _fDemandEff > _fReadyCap THEN
        _bGap := TRUE;                      // 供气缺口（信息级，不超载投切） / Supply gap, no overload dispatch
        _fDemandEff := _fReadyCap;          // 投切按就绪池全量封顶（安全侧） / Dispatch capped at the ready pool
    END_IF
    _fSupplyCap := 0.0;                     // 投运池能力清零 / Dispatched capacity cleared
    _uNeed := 0;                            // 需投台数清零 / Units needed cleared
    FOR _uIdx := 1 TO DL_UNIT_MAX DO
        IF _uIdx <= DL_UNIT_MAX THEN        // 二次闸 / Secondary gate
            IF abUnitReady[_uIdx] AND (NOT _abUnitBanned[_uIdx])
               AND (_fSupplyCap < _fDemandEff) THEN
                abUnitCmd[_uIdx] := TRUE;   // 投运指令置位 / Dispatch command set
                IF (aN2SupplyNm3H[_uIdx] <> aN2SupplyNm3H[_uIdx]) OR (ABS(aN2SupplyNm3H[_uIdx]) > DL_AC_INF) THEN
                    (* 非有限能力台不参与累加（段 4 已剔除，此处双保险） / Non-finite excluded, double-guarded *)
                    _fSupplyCap := _fSupplyCap + 0.0; // 零贡献 / Zero contribution
                ELSE
                    _fSupplyCap := _fSupplyCap + aN2SupplyNm3H[_uIdx]; // 投运能力累加 / Dispatched capacity accumulated
                END_IF
                _uNeed := _uNeed + 1;       // 需投台数递增 / Units needed increment
            END_IF
        END_IF
    END_FOR
    uUnitsNeeded := _uNeed;                 // 需投台数出口 / Units needed outlet
    fSupplyMarginNm3H := _fReadyCap - fN2DemandNm3H; // 余量出口（负值即缺口，按原始需求算） / Margin outlet, negative means a gap
END_IF

(*------------------------------------------------------------------------------
 * 段 6｜各台启动反馈确认计时无条件刷新（R40：CASE 之外每拍必调）
 *      Per-unit feedback timers refreshed unconditionally per R40
 *-----------------------------------------------------------------------------*)
FOR _uIdx := 1 TO DL_UNIT_MAX DO
    IF _uIdx <= DL_UNIT_MAX THEN            // 二次闸 / Secondary gate
        aFbDelay[_uIdx](IN := abUnitCmd[_uIdx] AND (NOT abUnitRunFb[_uIdx]) AND (NOT _aFbBreak[_uIdx]),
                        PT := tStartFbDelay); // 启动反馈确认计时 / Start-feedback confirm timer
        _aFbBreak[_uIdx] := FALSE;          // 断输入拍在调用后自清 / Break self-cleared after the call
        IF aFbDelay[_uIdx].Q THEN
            _abUnitBanned[_uIdx] := TRUE;   // 启动失败：剔除轮值池 / Start failure, unit banned
            _bAnyBanned := TRUE;            // 剔除标志置位 / Banned flag raised
            _aFbBreak[_uIdx] := TRUE;       // 窗重启（下次投切重新计时） / The window restarts for the next dispatch
        END_IF
    END_IF
END_FOR

(*------------------------------------------------------------------------------
 * 段 7｜码位出口
 *      Code outlet
 *-----------------------------------------------------------------------------*)
IF _bIllegal THEN
    eErr   := 16#0005_0326;                 // 故障级：状态机兜底 / Fault: fallback
    bError := TRUE;                         // 置故障标志 / Raise the fault flag
ELSIF _bDemandBad OR _bAnyBanned THEN
    eErr   := 16#0005_0324;                 // 故障级：启动失败/非有限剔除（R90 复用） / Fault: start failure or non-finite ban
    bError := TRUE;                         // 置故障标志 / Raise the fault flag
    bValid := TRUE;                         // 调度结果本身可用（剔除台已隔离） / The dispatch result itself is usable
ELSIF _bGap THEN
    eErr := 16#0005_01EA;                   // 信息级：供气缺口（不超载投切） / Info: supply gap, no overload dispatch
    bValid := TRUE;                         // 输出可用 / Outputs usable
ELSE
    bValid := bEnable;                      // 使能且正常：输出可用 / Outputs usable when enabled
END_IF
END_FUNCTION_BLOCK

(* ---- FB_DL_AirCompressorMasterSeq.st ---- *)
(*
  Name: FB_DL_AirCompressorMasterSeq
  Category: DL_Process
  Version: 1.0.0
  Round: R90 / 2026-11-25
  开源溯源：clean-room 自研（族 压缩空气系统能效，ST 开源生态实测 0 命中，无外部代码引入）
  功能：1) 两机空压站群控：主用机常开承担基载，压力跌破加载点且单机不够时投入辅机（双机运行），
           压力回到卸载点以上则退出辅机，回到单机主用相，形成带迟滞的两级容量控制。
        2) 主备轮换：主用相由轮换定时器 tonRot 计时（PT = tRotateH），到点后比较两机累计运行小时，
           把小时较少的一台设为主用，实现运行小时均衡；定时器自复位（IN := 运行相 AND NOT Q），
           不依赖外部沿清零。
        3) 故障切换：主用机故障立即由备机接管（相位在主用相之间直接迁移，不落故障相）；
           仅在两台同时故障或组态非法时才进故障相并锁存码值。辅机故障则退回单机主用相。
        4) 加载/卸载由带回差的锁存量给出：压力 <= 加载点置加载锁存，>= 卸载点清加载锁存，
           带内保持，防止在压力带内高频加减载。
  边界条件：1) 非有限值闸：压力、目标、回差、扫描周期四路实值入参统一过
           NOT(x > -DL_BIG AND x < DL_BIG)，同时拦 NaN 与 Inf；命中即判组态非法并进故障相，
           绝不把 NaN 送进压力比较（NaN 比较恒假会让加载判据静默失效，R19）。
        2) 组态零闸：fTargetBar 必须 > DL_EPS；fHystBar 必须 >= DL_HYST_MIN 且 <= fTargetBar
           （回差为 0 或越界会使加载点 >= 卸载点，压力带反号或退化为单点，必然频繁启停）；
           ABS(fCycleS) > DL_EPS 才允许累计运行小时（R21：斜率/积分类算法必须把周期时间作为入参
           并做零闸，不许假设固定扫描周期）。
        3) 压力带钳制：fTargetBar 钳 0 ~ DL_P_MAX(40 bar)、fHystBar 钳 0 ~ DL_P_MAX，
           加载点再钳到 >= 0，卸载点钳到 <= DL_P_MAX，防组态越界把压力带推到量程外。
        4) 饱和钳制：累计运行小时钳 0 ~ DL_H_MAX(200000 h)，防长年运行溢出。
        5) 相超时说明：eAcmLead1/eAcmLead2 两相的「超时」由轮换定时器 tonRot 承担（到点即轮换，
           该定时器本身就是主用相的时限监视）；eAcmAssist1/eAcmAssist2 两相由 tonAssist 监视
           （投入辅机后 DL_ASSIST_MAX 内压力仍未恢复 → 气量不足，判故障）；
           eAcmIdle 与 eAcmFault 为稳态相等候相，不设超时（设了会周期性误报）。
        6) 状态机兜底：CASE 全态覆盖 + ELSE 强制回故障相；故障解除路径为
           (NOT xAuto) AND (NOT xFault1) AND (NOT xFault2)，可达。
        7) FB 主体不使用 RETURN，统一单出口（跨平台可移植性）。
  量纲自证：fLoadBar = bar − bar/2 = bar；fUnloadBar = bar + bar/2 = bar；
           运行小时 = (s) / (s/h) = h，与 fHours1/fHours2 同量纲；
           tonRot/tonAssist 的 PT 为 [TIME]，与 TON 同量纲；本件无跨量纲相加。
  码表 Error codes（本件格 0090_04xx，故障级一律 3 行内置 _uFault/_bFault/_eState）:
    16#0090_0401 信息级：自动未投入（不置故障位）
    16#0090_0402 故障级：两台空压机同时故障
    16#0090_0403 故障级：辅机投入后压力长时间未恢复（气量不足）
    16#0090_0404 故障级：组态非法（目标压力/回差/扫描周期越界或非有限）
    16#0090_0405 故障级：状态机落 ELSE 兜底（非法相位 ID）

  修订历史 Revision :
    2026-11-25  v1.0.0  R90 首版
*)

TYPE E_DL_AcmState :
(
    eAcmIdle    := 0,    // 待机：自动未投入 / Idle, automatic mode not engaged
    eAcmLead1   := 10,   // 1 号主用，2 号停机 / Unit 1 lead, unit 2 stopped
    eAcmLead2   := 20,   // 2 号主用，1 号停机 / Unit 2 lead, unit 1 stopped
    eAcmAssist1 := 30,   // 1 号为主 + 2 号辅，双机运行 / Unit 1 lead with unit 2 assisting
    eAcmAssist2 := 40,   // 2 号为主 + 1 号辅，双机运行 / Unit 2 lead with unit 1 assisting
    eAcmFault   := 90    // 故障：锁存待解除 / Fault, latched awaiting release
);
END_TYPE

FUNCTION_BLOCK FB_DL_AirCompressorMasterSeq
VAR_INPUT
    xAuto        : BOOL;    // 自动投入指令 [bool] / Automatic mode command [bool]
    xFault1      : BOOL;    // 1 号机故障汇总 [bool] / Unit 1 fault aggregate [bool]
    xFault2      : BOOL;    // 2 号机故障汇总 [bool] / Unit 2 fault aggregate [bool]
    fPressureBar : REAL;    // 母管压力实测 [bar] / Header pressure measurement [bar]
    fTargetBar   : REAL;    // 目标压力（压力带中心）[bar] / Target pressure, band centre [bar]
    fHystBar     : REAL;    // 加载/卸载回差带宽 [bar] / Load-unload hysteresis band [bar]
    tRotateH     : TIME;    // 主备轮换周期 [TIME] / Lead rotation period [TIME]
    fCycleS      : REAL;    // 扫描周期 [s] / Scan cycle time [s]
END_VAR
VAR_OUTPUT
    xRun1        : BOOL;    // 1 号机运行指令 [bool] / Unit 1 run command [bool]
    xRun2        : BOOL;    // 2 号机运行指令 [bool] / Unit 2 run command [bool]
    xLoad1       : BOOL;    // 1 号机加载指令 [bool] / Unit 1 load command [bool]
    xLoad2       : BOOL;    // 2 号机加载指令 [bool] / Unit 2 load command [bool]
    fLoadBar     : REAL;    // 加载压力点 [bar] / Load pressure point [bar]
    fUnloadBar   : REAL;    // 卸载压力点 [bar] / Unload pressure point [bar]
    fHours1      : REAL;    // 1 号机累计运行小时 [h] / Unit 1 accumulated running hours [h]
    fHours2      : REAL;    // 2 号机累计运行小时 [h] / Unit 2 accumulated running hours [h]
    eState       : E_DL_AcmState;   // 状态出口，段尾单点映射 / State outlet, single-point mapped
    nErrId       : UDINT;   // 事件码，0 = 无事件 / Event code, 0 = none
END_VAR
VAR
    tonRot       : TON;     // 主用相轮换定时器，自复位 [TIME] / Lead rotation timer, self-resetting
    tonAssist    : TON;     // 辅机投入恢复监视定时器 [TIME] / Assist recovery supervision timer
    _eState      : E_DL_AcmState := E_DL_AcmState.eAcmIdle;   // 内部相位（CASE 唯一写入目标）
    _eStatePrev  : E_DL_AcmState := E_DL_AcmState.eAcmIdle;   // 上一拍相位快照（周期末更新）
    _fTargetClamp: REAL;    // 钳制后的目标压力 [bar] / Clamped target pressure [bar]
    _fHystClamp  : REAL;    // 钳制后的回差带宽 [bar] / Clamped hysteresis band [bar]
    _fLoadPtBar  : REAL;    // 加载压力点 [bar] / Load pressure point [bar]
    _fUnloadPtBar: REAL;    // 卸载压力点 [bar] / Unload pressure point [bar]
    _bNeedAssist : BOOL;    // 需投入辅机（压力跌破加载点）[bool] / Assist required flag [bool]
    _bRecovered  : BOOL;    // 压力已回到卸载点以上 [bool] / Pressure recovered flag [bool]
    _bLeadRunning: BOOL;    // 主用相运行中（轮换定时器激励源）[bool] / Lead phase running flag [bool]
    _bRun1       : BOOL;    // 1 号机运行内部量 [bool] / Unit 1 run internal [bool]
    _bRun2       : BOOL;    // 2 号机运行内部量 [bool] / Unit 2 run internal [bool]
    _bLoadLat1   : BOOL;    // 1 号机加载锁存（迟滞承载）[bool] / Unit 1 load latch [bool]
    _bLoadLat2   : BOOL;    // 2 号机加载锁存（迟滞承载）[bool] / Unit 2 load latch [bool]
    _fHours1     : REAL;    // 1 号机累计运行小时内部量 [h] / Unit 1 hours internal [h]
    _fHours2     : REAL;    // 2 号机累计运行小时内部量 [h] / Unit 2 hours internal [h]
    _bCfgBad     : BOOL;    // 组态非法聚合 [bool] / Configuration invalid aggregate [bool]
    _bFault      : BOOL;    // 故障锁存位 [bool] / Latched fault flag [bool]
    _uInfo       : UDINT;   // 信息码，每拍重算 / Info code, recomputed every cycle
    _uFault      : UDINT;   // 故障码锁存 / Latched fault code
END_VAR
VAR CONSTANT
    DL_EPS       : REAL := 1.0E-9;      // 组态零闸阈值 [-] / Configuration zero gate threshold [-]
    DL_BIG       : REAL := 1.0E12;      // 非有限值闸量级上限 [-] / Finiteness gate magnitude [-]
    DL_P_MAX     : REAL := 40.0;        // 压力量程上限 [bar] / Pressure range ceiling [bar]
    DL_HYST_MIN  : REAL := 0.05;        // 回差带宽下限 [bar] / Hysteresis lower bound [bar]
    DL_TWO       : REAL := 2.0;         // 半带宽除数（对称展开）[-] / Half-band divisor [-]
    DL_S_PER_H   : REAL := 3600.0;      // h → s 换算因子 [s/h] / Hour to second factor [s/h]
    DL_H_MAX     : REAL := 200000.0;    // 累计运行小时饱和上限 [h] / Running hours saturation ceiling [h]
    DL_ASSIST_MAX: TIME := T#30M;       // 辅机投入后压力恢复监视窗 [TIME] / Assist recovery window [TIME]
END_VAR

(* —— 段 0：单拍量预清零（锁存量 _uFault/_bFault/_bLoadLat*/_fHours*/_eStatePrev 不入清单，R187①） —— *)
_uInfo := 16#0090_0401;                     // 缺省信息：自动未投入（进自动后由各相覆盖）
nErrId := 16#0000_0000;                     // 事件码缺省无事件 / Event code defaults to none

(* —— 段 1：非有限值闸（R19：NaN 比较恒假会让加载判据静默失效，必须前置拦截） —— *)
_bCfgBad := NOT (fPressureBar > -DL_BIG AND fPressureBar < DL_BIG)
            OR NOT (fTargetBar > -DL_BIG AND fTargetBar < DL_BIG)
            OR NOT (fHystBar > -DL_BIG AND fHystBar < DL_BIG)
            OR NOT (fCycleS > -DL_BIG AND fCycleS < DL_BIG);

(* —— 段 2：组态零闸（R4/R21：回差退化、目标为零、周期为零均判组态非法） —— *)
_bCfgBad := _bCfgBad
            OR (fTargetBar <= DL_EPS)                         // 目标压力必须为正
            OR (fTargetBar > DL_P_MAX)                        // 目标压力不越量程
            OR (fHystBar < DL_HYST_MIN)                       // 回差不得低于下限（防频繁启停）
            OR (fHystBar > fTargetBar)                        // 回差不得大于目标压力（否则加载点为负）
            OR (ABS(fCycleS) <= DL_EPS);                      // 扫描周期零闸

(* —— 段 3：压力带解算（R22 方向自核：加载在下、卸载在上，各偏半个回差） —— *)
_fTargetClamp := LIMIT(0.0, fTargetBar, DL_P_MAX);            // 目标压力钳 0..40 [bar]
_fHystClamp := LIMIT(0.0, fHystBar, DL_P_MAX);                // 回差钳 0..40 [bar]
_fLoadPtBar := LIMIT(0.0, _fTargetClamp - _fHystClamp / DL_TWO, DL_P_MAX);      // 加载点 [bar]
_fUnloadPtBar := LIMIT(0.0, _fTargetClamp + _fHystClamp / DL_TWO, DL_P_MAX);    // 卸载点 [bar]

(* —— 段 4：判据量（压力越低越需辅机，回到卸载点以上即判恢复） —— *)
_bNeedAssist := (NOT _bCfgBad) AND (fPressureBar <= _fLoadPtBar);      // 跌破加载点
_bRecovered := (NOT _bCfgBad) AND (fPressureBar >= _fUnloadPtBar);     // 回到卸载点以上

(* —— 段 5：定时器无条件周期刷新（R7 + R188：轮换定时器自复位，不靠外部沿） —— *)
_bLeadRunning := (_eState = E_DL_AcmState.eAcmLead1) OR (_eState = E_DL_AcmState.eAcmLead2);
tonRot(IN := _bLeadRunning AND (NOT tonRot.Q), PT := tRotateH);        // 主用相轮换计时，自复位
tonAssist(IN := (_eState = E_DL_AcmState.eAcmAssist1) OR (_eState = E_DL_AcmState.eAcmAssist2),
          PT := DL_ASSIST_MAX);                                        // 辅机恢复监视窗

(* —— 段 6：全局故障拦截（优先级最高；已锁存则不再改写码值，禁同拍抹除） —— *)
IF _bCfgBad AND (NOT _bFault) THEN
    _uFault := 16#0090_0404;                // 故障级：组态非法
    _bFault := TRUE;                        // 锁存（3 行内置，R45 配对）
    _eState := E_DL_AcmState.eAcmFault;
END_IF
IF xFault1 AND xFault2 AND (NOT _bFault) THEN
    _uFault := 16#0090_0402;                // 故障级：两机同时故障
    _bFault := TRUE;                        // 锁存
    _eState := E_DL_AcmState.eAcmFault;
END_IF

(* —— 段 7：相位机（只做迁移；出口在段 9 单点映射） —— *)
CASE _eState OF

E_DL_AcmState.eAcmIdle:
    IF NOT xAuto THEN
        _uInfo := 16#0090_0401;             // 信息级：自动未投入
    ELSIF _fHours1 <= _fHours2 THEN
        _eState := E_DL_AcmState.eAcmLead1; // 小时较少者为主用（均衡起点）
    ELSE
        _eState := E_DL_AcmState.eAcmLead2;
    END_IF

E_DL_AcmState.eAcmLead1:
    IF NOT xAuto THEN
        _eState := E_DL_AcmState.eAcmIdle;  // 撤自动：回待机
    ELSIF xFault1 THEN
        _eState := E_DL_AcmState.eAcmLead2; // 主用故障：备机接管（不落故障相）
    ELSIF _bNeedAssist THEN
        _eState := E_DL_AcmState.eAcmAssist1;   // 单机不足：投入辅机
    ELSIF tonRot.Q AND (_fHours2 < _fHours1) THEN
        _eState := E_DL_AcmState.eAcmLead2; // 轮换到点且 2 号小时更少：换主用
    END_IF

E_DL_AcmState.eAcmLead2:
    IF NOT xAuto THEN
        _eState := E_DL_AcmState.eAcmIdle;
    ELSIF xFault2 THEN
        _eState := E_DL_AcmState.eAcmLead1; // 主用故障：备机接管
    ELSIF _bNeedAssist THEN
        _eState := E_DL_AcmState.eAcmAssist2;
    ELSIF tonRot.Q AND (_fHours1 < _fHours2) THEN
        _eState := E_DL_AcmState.eAcmLead1; // 轮换到点且 1 号小时更少：换主用
    END_IF

E_DL_AcmState.eAcmAssist1:
    IF NOT xAuto THEN
        _eState := E_DL_AcmState.eAcmIdle;
    ELSIF xFault1 THEN
        _eState := E_DL_AcmState.eAcmLead2; // 主机故障：辅机转主用
    ELSIF xFault2 THEN
        _eState := E_DL_AcmState.eAcmLead1; // 辅机故障：退回单机主用
    ELSIF _bRecovered THEN
        _eState := E_DL_AcmState.eAcmLead1; // 本拍合法事件（压力恢复）优先于超时迁移（R275）
    ELSIF tonAssist.Q THEN
        _uFault := 16#0090_0403;            // 故障级：气量不足，双机仍不能恢复压力
        _bFault := TRUE;
        _eState := E_DL_AcmState.eAcmFault;
    END_IF

E_DL_AcmState.eAcmAssist2:
    IF NOT xAuto THEN
        _eState := E_DL_AcmState.eAcmIdle;
    ELSIF xFault2 THEN
        _eState := E_DL_AcmState.eAcmLead1; // 主机故障：辅机转主用
    ELSIF xFault1 THEN
        _eState := E_DL_AcmState.eAcmLead2; // 辅机故障：退回单机主用
    ELSIF _bRecovered THEN
        _eState := E_DL_AcmState.eAcmLead2; // 本拍合法事件优先于超时迁移
    ELSIF tonAssist.Q THEN
        _uFault := 16#0090_0403;            // 故障级：气量不足
        _bFault := TRUE;
        _eState := E_DL_AcmState.eAcmFault;
    END_IF

E_DL_AcmState.eAcmFault:
    IF (NOT xAuto) AND (NOT xFault1) AND (NOT xFault2) AND (NOT _bCfgBad) THEN
        _bFault := FALSE;                   // 解除路径：撤自动 + 两机故障消失 + 组态恢复（可达）
        _uFault := 16#0000_0000;            // 清锁存码
        _eState := E_DL_AcmState.eAcmIdle;  // 回待机
    END_IF

ELSE
    _uFault := 16#0090_0405;                // 故障级：非法相位 ID 兜底
    _bFault := TRUE;                        // 锁存
    _eState := E_DL_AcmState.eAcmFault;     // 强制回故障相

END_CASE

(* —— 段 8：后置段（R23：运行派生、加载锁存、小时累计一律在迁移判断之后） —— *)
_bRun1 := ((_eState = E_DL_AcmState.eAcmLead1) OR (_eState = E_DL_AcmState.eAcmAssist1)
           OR (_eState = E_DL_AcmState.eAcmAssist2)) AND (NOT _bFault) AND (NOT xFault1);
_bRun2 := ((_eState = E_DL_AcmState.eAcmLead2) OR (_eState = E_DL_AcmState.eAcmAssist1)
           OR (_eState = E_DL_AcmState.eAcmAssist2)) AND (NOT _bFault) AND (NOT xFault2);

(* 加载锁存：跌破加载点置位，回到卸载点以上复位，带内保持（迟滞防频繁加减载） *)
IF NOT _bRun1 THEN
    _bLoadLat1 := FALSE;                    // 停机即清加载锁存
ELSIF fPressureBar <= _fLoadPtBar THEN
    _bLoadLat1 := TRUE;                     // 跌破加载点：加载
ELSIF fPressureBar >= _fUnloadPtBar THEN
    _bLoadLat1 := FALSE;                    // 回到卸载点以上：卸载
END_IF
IF NOT _bRun2 THEN
    _bLoadLat2 := FALSE;                    // 停机即清加载锁存
ELSIF fPressureBar <= _fLoadPtBar THEN
    _bLoadLat2 := TRUE;                     // 跌破加载点：加载
ELSIF fPressureBar >= _fUnloadPtBar THEN
    _bLoadLat2 := FALSE;                    // 回到卸载点以上：卸载
END_IF

(* 运行小时累计（R21：周期时间已做零闸，段 2 已判 ABS(fCycleS) > DL_EPS 才允许进入本段） *)
IF _bRun1 AND (ABS(fCycleS) > DL_EPS) THEN
    _fHours1 := MIN(DL_H_MAX, _fHours1 + fCycleS / DL_S_PER_H);    // s / (s/h) = h
END_IF
IF _bRun2 AND (ABS(fCycleS) > DL_EPS) THEN
    _fHours2 := MIN(DL_H_MAX, _fHours2 + fCycleS / DL_S_PER_H);    // s / (s/h) = h
END_IF

_eStatePrev := _eState;                     // 快照统一在周期末尾更新（R23）

(* —— 段 9：出口单点映射（名实同源；运行/加载由状态与锁存导出，不在多分支各写一遍） —— *)
xRun1 := _bRun1;                            // 1 号机运行出口
xRun2 := _bRun2;                            // 2 号机运行出口
xLoad1 := _bRun1 AND _bLoadLat1;            // 1 号机加载出口（停机必不加载）
xLoad2 := _bRun2 AND _bLoadLat2;            // 2 号机加载出口
IF _bCfgBad THEN
    fLoadBar := 0.0;                        // 组态非法：压力带出口闸断为字面量，禁 NaN 外泄
    fUnloadBar := 0.0;                      // 同上
ELSIF _bFault THEN
    fLoadBar := _fLoadPtBar;                // 故障锁存但组态仍有效：回放上拍解算值
    fUnloadBar := _fUnloadPtBar;            // 同上
ELSE
    fLoadBar := _fLoadPtBar;                // 加载压力点出口 [bar]
    fUnloadBar := _fUnloadPtBar;            // 卸载压力点出口 [bar]
END_IF
fHours1 := _fHours1;                        // 1 号机运行小时出口 [h]
fHours2 := _fHours2;                        // 2 号机运行小时出口 [h]
eState := _eState;                          // 状态出口单点映射
IF _bFault THEN
    nErrId := _uFault;                      // 故障锁存码回放（不在故障相按当下输入重推断）
ELSE
    nErrId := _uInfo;                       // 信息码
END_IF

END_FUNCTION_BLOCK

(* ---- FB_DL_AirLeakDecayTest.st ---- *)
(*
  组件名 Component   : FB_DL_AirLeakDecayTest
  子库 Sublibrary    : DL_Process
  版本 Version       : 1.0.0
  兼容性 Platform    : CODESYS 3.5 / TwinCAT 3 / 汇川 InoProShop / Machine Expert（仅 Standard.library）
  功能 Function      : 气密压降法泄漏测试（与 FC 氦检分工：空气压降 vs 氦质谱）：
                       1) 三段顺控：充压（eCharge，出充压指令至测试压力确认）→
                       稳压（eStabilize，驻留 tStabDur 待温度平衡）→ 测量（eMeasure，
                       驻留 tMeasDur，窗始/窗末压力双快照）；
                       2) 温度补偿：绝对温标折算，压降补偿值 =
                       p1 - p2 × (T1/T2)，T 为绝对温度（摄氏度 + 开尔文偏置）；
                       3) 泄漏率换算判级：泄漏率 = 补偿压降 × 容积 / 测量时长，
                       <= fLeakLim 判合格，否则不合格；
                       4) 测量段压力跌破 fPressMinPa → 充压丢失故障锁存。
  边界 Boundary      : ① 本件只出充压指令与测试结论，不写物理 IO；
                       ② 除法前置域闸：测量时长秒值下限 1.0 s、绝对温度下限
                       1.0 K、容积 > 0（组态闸承载）；
                       ③ 各相计时独立 TON 实例（禁跨相复用）；窗始快照进相首拍
                       写定，锁存回放不重扫；
                       ④ 故障锁存解除唯一路径 = bReset 上升沿（输入引脚，恒可达）；
                       ⑤ 无全局变量引用、无外部变量声明、无物理地址寻址。
  依赖 Depends       : Standard.library（R_TRIG / TON）
  溯源 Origin        : 道莅自研 clean-room（自研行业池：通用质量工装气密检测
                       共性语义，零外部代码行复制）
  码位 Code          : 16#06_0_C2（Process 段 0006，C 子带 C2 格）
  码表 Error codes（本件格 06_0_C2，单轨子道：故障 0x02C2 / 信息 0x01C2）:
    16#0006_02C2 故障级：气密测试故障总码（充压超时 / 测量段压力跌破下限 /
                 组态非法 / 输入非有限），锁存至复位
    16#0006_01C2 信息级：测试结论写定沿（合格或不合格判定拍）
  修订历史 Revision  :
    2026-11-19  v1.0.0  R44 首版（批次 4 · 序号 19）
*)

TYPE E_DL_AltPhase :
(
    eIdle      := 0,   // 空闲：等测试沿 / Idle, waiting test edge
    eCharge    := 10,  // 充压：至测试压力确认 / Charging to test pressure
    eStabilize := 20,  // 稳压：温度平衡驻留 / Stabilizing dwell
    eMeasure   := 30,  // 测量：双快照驻留 / Measuring dwell
    eDone      := 40,  // 完成：结论驻留 / Done, verdict held
    eFault     := 90   // 故障：总码锁存 / Fault, latched
);
END_TYPE

FUNCTION_BLOCK FB_DL_AirLeakDecayTest
VAR_INPUT
    bEnable      : BOOL;                   // 使能（电平）[-] / Enable
    bReset       : BOOL;                   // 上升沿清故障锁存 [-] / Reset edge
    bTestCmd     : BOOL;                   // 测试指令（上升沿承载）[-] / Test command edge
    fPressPa     : REAL;                   // 腔体实测压力 [帕斯卡] / Measured pressure
    fTempC       : REAL;                   // 腔体实测温度 [摄氏度] / Measured temperature
    fTestPressPa : REAL := 500000.0;       // 测试压力 [帕斯卡] / Test pressure
    fPressMinPa  : REAL := 400000.0;       // 测量段压力下限 [帕斯卡] / Measurement pressure floor
    fVolumeL     : REAL := 10.0;           // 腔体容积 [升] / Cavity volume
    fLeakLimPaLs : REAL := 1.0;            // 泄漏率合格限 [帕·升/秒] / Leak rate pass limit
    tStabDur     : TIME := T#60S;          // 稳压驻留 [毫秒] / Stabilization dwell
    tMeasDur     : TIME := T#120S;         // 测量驻留 [毫秒] / Measurement dwell
    tChargeTo    : TIME := T#120S;         // 充压超时 [毫秒] / Charge timeout
END_VAR
VAR_OUTPUT
    bChargeCmd   : BOOL;                   // 充压指令输出 [-] / Charge command output
    bTestPass    : BOOL;                   // 结论：合格 [-] / Verdict pass flag
    fLeakRatePaLs: REAL;                   // 实测泄漏率 [帕·升/秒] / Measured leak rate
    fDpCompPa    : REAL;                   // 温度补偿压降 [帕斯卡] / Compensated pressure drop
    ePhase       : E_DL_AltPhase;          // 相位出口，段尾单点映射 / Phase outlet
    bError       : BOOL;                   // 故障锁存标志 [-] / Fault latch flag
    uErrId       : UDINT;                  // 事件码，0 = 无事件 / Event code
END_VAR
VAR
    rtReset: R_TRIG;                       // 复位沿实例，段 0 无条件刷新 / Reset edge
    rtTest : R_TRIG;                       // 测试沿实例，段 0 无条件刷新 / Test edge
    tonStabDur: TON;                       // 稳压驻留计时（独立实例） / Stabilization timer
    tonMeasDur: TON;                       // 测量驻留计时（独立实例） / Measurement timer
    tonChargeTo: TON;                      // 充压超时（专用超时件命名） / Charge timeout
    _ePhase: E_DL_AltPhase := E_DL_AltPhase.eIdle;     // 内部相位（CASE 唯一写入目标）/ Internal phase
    _fP1Pa : REAL;                         // 窗始压力快照 [帕斯卡] / Window-start pressure snapshot
    _fT1C  : REAL;                         // 窗始温度快照 [摄氏度] / Window-start temperature snapshot
    _bSnapDone: BOOL;                      // 窗始快照已取标志 [-] / Snapshot taken flag
    _fT1K  : REAL;                         // 窗始绝对温度 [开尔文] / Window-start absolute temperature
    _fT2K  : REAL;                         // 窗末绝对温度 [开尔文] / Window-end absolute temperature
    _bFault: BOOL;                         // 故障锁存位（锁存量） / Latched fault bit
    _uFault: UDINT;                        // 故障码锁存（锁存量） / Latched fault code
    _bCfgBad: BOOL;                        // 组态非法当拍量 [-] / Config illegal flag
    _bNonFin: BOOL;                        // 输入非有限当拍量 [-] / Non-finite input flag
END_VAR
VAR CONSTANT
    DL_KELVIN_OFF : REAL := 273.15;        // 开尔文偏置 [开尔文] / Kelvin offset
    DL_T_ABS_MIN  : REAL := 1.0;           // 绝对温度下限 [开尔文] / Absolute temperature floor
    DL_MEAS_MIN_S : REAL := 1.0;           // 测量时长秒值下限 [秒] / Measurement seconds floor
    DL_MS_PER_S   : REAL := 1000.0;        // 毫秒 → 秒换算系数 [毫秒/秒] / Milliseconds per second
    DL_ABS_MAX    : REAL := 1.0E30;        // 有限值判定上界 [工程单位] / Finite bound
    DL_ZERO       : REAL := 0.0;           // 零常量 [工程单位] / Zero constant
END_VAR

(* —— 段 0｜沿与定时器每拍无条件刷新（禁置于 IF/CASE 内；各相独立实例禁复用） —— *)
rtReset(CLK := bReset);
rtTest (CLK := bTestCmd);
tonStabDur (IN := (_ePhase = E_DL_AltPhase.eStabilize) AND (NOT _bFault), PT := tStabDur);
tonMeasDur (IN := (_ePhase = E_DL_AltPhase.eMeasure) AND (NOT _bFault), PT := tMeasDur);
tonChargeTo(IN := (_ePhase = E_DL_AltPhase.eCharge) AND (NOT _bFault), PT := tChargeTo);

(* —— 段 1｜瞬时量预清零（锁存量 _bFault/_uFault/bTestPass/_fP1Pa 不入清单） —— *)
uErrId   := 16#0000_0000;
_bCfgBad := FALSE;
_bNonFin := FALSE;

(* —— 段 2｜复位沿：故障一次性清干净，相位回空闲，充压指令撤销 —— *)
IF rtReset.Q THEN
    _bFault := FALSE;
    _uFault := 16#0000_0000;
    bChargeCmd := FALSE;
    _ePhase := E_DL_AltPhase.eIdle;
END_IF

(* —— 段 3｜组态闸与非有限判据（覆盖全部参与判据换算引脚） —— *)
IF (fTestPressPa <= fPressMinPa) OR (fPressMinPa <= DL_ZERO) OR (fVolumeL <= DL_ZERO)
   OR (fLeakLimPaLs <= DL_ZERO) OR (tStabDur = T#0S) OR (tMeasDur = T#0S)
   OR (tChargeTo = T#0S) THEN
    _bCfgBad := TRUE;
END_IF
IF (fPressPa <> fPressPa) OR ((fPressPa - fPressPa) <> DL_ZERO)
   OR (fTempC <> fTempC) OR ((fTempC - fTempC) <> DL_ZERO) THEN
    _bNonFin := TRUE;
END_IF

(* —— 段 4｜主状态机：六态全覆盖 + ELSE 兜底 —— *)
CASE _ePhase OF

E_DL_AltPhase.eIdle:
    bChargeCmd := FALSE;
    IF rtTest.Q AND bEnable AND (NOT _bFault) AND (NOT _bCfgBad) AND (NOT _bNonFin) THEN
        bTestPass := FALSE;
        fLeakRatePaLs := DL_ZERO;
        fDpCompPa := DL_ZERO;
        _bSnapDone := FALSE;
        _ePhase := E_DL_AltPhase.eCharge;
    ELSIF rtTest.Q AND (_bFault OR _bCfgBad OR _bNonFin) THEN
        _bFault := TRUE;                 // 带病启动拒绝
        _uFault := 16#0006_02C2;
        bError  := TRUE;
        _ePhase := E_DL_AltPhase.eFault;
    END_IF

E_DL_AltPhase.eCharge:
    bChargeCmd := TRUE;
    IF _bNonFin THEN
        _bFault := TRUE;
        _uFault := 16#0006_02C2;
        bError  := TRUE;
        _ePhase := E_DL_AltPhase.eFault;
    ELSIF fPressPa >= fTestPressPa THEN
        bChargeCmd := FALSE;
        _ePhase := E_DL_AltPhase.eStabilize;     // 迁出条件 1：测试压力达成
    ELSIF tonChargeTo.Q THEN
        _bFault := TRUE;                 // 迁出条件 2（故障路）：充压超时
        _uFault := 16#0006_02C2;
        bError  := TRUE;
        bChargeCmd := FALSE;
        _ePhase := E_DL_AltPhase.eFault;
    END_IF

E_DL_AltPhase.eStabilize:
    bChargeCmd := FALSE;
    IF _bNonFin THEN
        _bFault := TRUE;
        _uFault := 16#0006_02C2;
        bError  := TRUE;
        _ePhase := E_DL_AltPhase.eFault;
    ELSIF tonStabDur.Q THEN
        _bSnapDone := FALSE;
        _ePhase := E_DL_AltPhase.eMeasure;   // 稳压驻留完成：进测量相
    END_IF

E_DL_AltPhase.eMeasure:
    bChargeCmd := FALSE;
    IF _bNonFin THEN
        _bFault := TRUE;
        _uFault := 16#0006_02C2;
        bError  := TRUE;
        _ePhase := E_DL_AltPhase.eFault;
    ELSIF fPressPa < fPressMinPa THEN
        _bFault := TRUE;                 // 测量段压力跌破下限：充压丢失
        _uFault := 16#0006_02C2;
        bError  := TRUE;
        _ePhase := E_DL_AltPhase.eFault;
    ELSIF NOT _bSnapDone THEN
        _fP1Pa := fPressPa;              // 窗始双快照：进相首拍写定（锁存回放不重扫）
        _fT1C  := fTempC;
        _bSnapDone := TRUE;
    ELSIF tonMeasDur.Q THEN
        (* 温度补偿判级：绝对温标折算，除子 = 绝对温度/测量时长，域闸均已过 *)
        _fT1K := _fT1C + DL_KELVIN_OFF;
        _fT2K := fTempC + DL_KELVIN_OFF;
        IF (_fT1K >= DL_T_ABS_MIN) AND (_fT2K >= DL_T_ABS_MIN) THEN
            fDpCompPa := _fP1Pa - (fPressPa * _fT1K / _fT2K);   // 补偿压降
            fLeakRatePaLs := MAX(fDpCompPa, DL_ZERO) * fVolumeL
                             / MAX(TIME_TO_REAL(tMeasDur) / DL_MS_PER_S, DL_MEAS_MIN_S);
            bTestPass := fLeakRatePaLs <= fLeakLimPaLs;
            uErrId := 16#0006_01C2;      // 信息级：结论写定沿
            _ePhase := E_DL_AltPhase.eDone;
        ELSE
            _bFault := TRUE;             // 绝对温度越下限：判据不可信
            _uFault := 16#0006_02C2;
            bError  := TRUE;
            _ePhase := E_DL_AltPhase.eFault;
        END_IF
    END_IF

E_DL_AltPhase.eDone:
    bChargeCmd := FALSE;
    IF NOT bTestCmd THEN
        _ePhase := E_DL_AltPhase.eIdle;  // 测试指令撤销：回空闲（结论锁存保留）
    END_IF

E_DL_AltPhase.eFault:
    bChargeCmd := FALSE;                 // 故障相：充压指令安全侧撤销
    bError := TRUE;
    ;                                    // 故障相驻留：只认复位沿（段 2 迁出）

ELSE
    _bFault := TRUE;                     // 兜底：非法相位锁存
    _uFault := 16#0006_02C2;
    bError  := TRUE;
    _ePhase := E_DL_AltPhase.eFault;
END_CASE

(* —— 段 5｜相位出口单点映射 —— *)
ePhase := _ePhase;
END_FUNCTION_BLOCK
